(* IEC 61131-3 sources: plc-st-coding-agent/progress/evidence/f14_v14_remaining_20261113/jobs/codex_minimax-m27, 165 files *)

(* ---- public-easy-01.candidate_01.st ---- *)
(* ENGINEERING_CONTRACT *)
(*
  State machine for bottle filling line with 6 sequential states:
  - IDLE (0): No outputs active. Waits for bottleSensor TRUE → CLEANING.
  - CLEANING (1): Pump_Motor active. cleaningConfirmButton TRUE → FILLING.
  - FILLING (2): Filling_Valve active. fillingConfirmButton TRUE → CAPPING.
  - CAPPING (3): Capping_Machine active. cappingConfirmButton TRUE → PACKAGING.
  - PACKAGING (4): Packing_Machine active. packingConfirmButton TRUE → COMPLETED.
  - COMPLETED (5): Completion_Light active (retention). finishedButton TRUE → IDLE.

  Outputs: Pump_Motor(FILLING), Filling_Valve(FILLING), Capping_Machine(CAPPING),
           Packing_Machine(PACKAGING), Completion_Light(COMPLETED,hold_until_reset).
  Reset: finishedButton deactivates Completion_Light and returns to IDLE.
*)
(* CONTRACT_RULES [* kind=hold_until_reset, output=Completion_Light, set_input=packingConfirmButton, reset_input=finishedButton *] *)

FUNCTION_BLOCK FillingLineControl
VAR
    currentState : INT := 0;
END_VAR

CASE currentState OF
    0: // IDLE
        Pump_Motor := FALSE;
        Filling_Valve := FALSE;
        Capping_Machine := FALSE;
        Packing_Machine := FALSE;
        Completion_Light := FALSE;

        IF bottleSensor THEN
            currentState := 1;
        END_IF;

    1: // CLEANING
        Pump_Motor := TRUE;
        Filling_Valve := FALSE;
        Capping_Machine := FALSE;
        Packing_Machine := FALSE;
        Completion_Light := FALSE;

        IF cleaningConfirmButton THEN
            currentState := 2;
        END_IF;

    2: // FILLING
        Pump_Motor := FALSE;
        Filling_Valve := TRUE;
        Capping_Machine := FALSE;
        Packing_Machine := FALSE;
        Completion_Light := FALSE;

        IF fillingConfirmButton THEN
            currentState := 3;
        END_IF;

    3: // CAPPING
        Pump_Motor := FALSE;
        Filling_Valve := FALSE;
        Capping_Machine := TRUE;
        Packing_Machine := FALSE;
        Completion_Light := FALSE;

        IF cappingConfirmButton THEN
            currentState := 4;
        END_IF;

    4: // PACKAGING
        Pump_Motor := FALSE;
        Filling_Valve := FALSE;
        Capping_Machine := FALSE;
        Packing_Machine := TRUE;
        Completion_Light := FALSE;

        IF packingConfirmButton THEN
            currentState := 5;
        END_IF;

    5: // COMPLETED
        Pump_Motor := FALSE;
        Filling_Valve := FALSE;
        Capping_Machine := FALSE;
        Packing_Machine := FALSE;
        Completion_Light := TRUE;

        IF finishedButton THEN
            currentState := 0;
        END_IF;
END_CASE;
END_FUNCTION_BLOCK

(* ---- public-easy-01.candidate_03.st ---- *)
(* ENGINEERING_CONTRACT *)
(*
  State machine for bottle filling line with 6 sequential states:
  - IDLE (0): No outputs active. Waits for bottleSensor TRUE → CLEANING.
  - CLEANING (1): Pump_Motor active. cleaningConfirmButton TRUE → FILLING.
  - FILLING (2): Filling_Valve active. fillingConfirmButton TRUE → CAPPING.
  - CAPPING (3): Capping_Machine active. cappingConfirmButton TRUE → PACKAGING.
  - PACKAGING (4): Packing_Machine active. packingConfirmButton TRUE → COMPLETED.
  - COMPLETED (5): Completion_Light active (retention). finishedButton TRUE → IDLE.

  Outputs: Pump_Motor(FILLING), Filling_Valve(FILLING), Capping_Machine(CAPPING),
           Packing_Machine(PACKAGING), Completion_Light(COMPLETED,hold_until_reset).
  Reset: finishedButton deactivates Completion_Light and returns to IDLE.
*)
(* CONTRACT_RULES [* kind=hold_until_reset, output=Completion_Light, set_input=packingConfirmButton, reset_input=finishedButton *] *)

FUNCTION_BLOCK FillingLineControl
VAR_INPUT
    bottleSensor : BOOL;
    cleaningConfirmButton : BOOL;
    fillingConfirmButton : BOOL;
    cappingConfirmButton : BOOL;
    packingConfirmButton : BOOL;
    finishedButton : BOOL;
END_VAR
VAR_OUTPUT
    Pump_Motor : BOOL;
    Filling_Valve : BOOL;
    Capping_Machine : BOOL;
    Packing_Machine : BOOL;
    Completion_Light : BOOL;
END_VAR
VAR
    currentState : INT := 0;
END_VAR

CASE currentState OF
    0: // IDLE
        Pump_Motor := FALSE;
        Filling_Valve := FALSE;
        Capping_Machine := FALSE;
        Packing_Machine := FALSE;
        Completion_Light := FALSE;

        IF bottleSensor THEN
            currentState := 1;
        END_IF;

    1: // CLEANING
        Pump_Motor := TRUE;
        Filling_Valve := FALSE;
        Capping_Machine := FALSE;
        Packing_Machine := FALSE;
        Completion_Light := FALSE;

        IF cleaningConfirmButton THEN
            currentState := 2;
        END_IF;

    2: // FILLING
        Pump_Motor := FALSE;
        Filling_Valve := TRUE;
        Capping_Machine := FALSE;
        Packing_Machine := FALSE;
        Completion_Light := FALSE;

        IF fillingConfirmButton THEN
            currentState := 3;
        END_IF;

    3: // CAPPING
        Pump_Motor := FALSE;
        Filling_Valve := FALSE;
        Capping_Machine := TRUE;
        Packing_Machine := FALSE;
        Completion_Light := FALSE;

        IF cappingConfirmButton THEN
            currentState := 4;
        END_IF;

    4: // PACKAGING
        Pump_Motor := FALSE;
        Filling_Valve := FALSE;
        Capping_Machine := FALSE;
        Packing_Machine := TRUE;
        Completion_Light := FALSE;

        IF packingConfirmButton THEN
            currentState := 5;
        END_IF;

    5: // COMPLETED
        Pump_Motor := FALSE;
        Filling_Valve := FALSE;
        Capping_Machine := FALSE;
        Packing_Machine := FALSE;
        Completion_Light := TRUE;

        IF finishedButton THEN
            currentState := 0;
        END_IF;
END_CASE;
END_FUNCTION_BLOCK

(* ---- public-easy-01.patch_base_02.st ---- *)
(* ENGINEERING_CONTRACT *)
(*
  State machine for bottle filling line with 6 sequential states:
  - IDLE (0): No outputs active. Waits for bottleSensor TRUE → CLEANING.
  - CLEANING (1): Pump_Motor active. cleaningConfirmButton TRUE → FILLING.
  - FILLING (2): Filling_Valve active. fillingConfirmButton TRUE → CAPPING.
  - CAPPING (3): Capping_Machine active. cappingConfirmButton TRUE → PACKAGING.
  - PACKAGING (4): Packing_Machine active. packingConfirmButton TRUE → COMPLETED.
  - COMPLETED (5): Completion_Light active (retention). finishedButton TRUE → IDLE.

  Outputs: Pump_Motor(FILLING), Filling_Valve(FILLING), Capping_Machine(CAPPING),
           Packing_Machine(PACKAGING), Completion_Light(COMPLETED,hold_until_reset).
  Reset: finishedButton deactivates Completion_Light and returns to IDLE.
*)
(* CONTRACT_RULES [* kind=hold_until_reset, output=Completion_Light, set_input=packingConfirmButton, reset_input=finishedButton *] *)

FUNCTION_BLOCK FillingLineControl
VAR
    currentState : INT := 0;
END_VAR

CASE currentState OF
    0: // IDLE
        Pump_Motor := FALSE;
        Filling_Valve := FALSE;
        Capping_Machine := FALSE;
        Packing_Machine := FALSE;
        Completion_Light := FALSE;

        IF bottleSensor THEN
            currentState := 1;
        END_IF;

    1: // CLEANING
        Pump_Motor := TRUE;
        Filling_Valve := FALSE;
        Capping_Machine := FALSE;
        Packing_Machine := FALSE;
        Completion_Light := FALSE;

        IF cleaningConfirmButton THEN
            currentState := 2;
        END_IF;

    2: // FILLING
        Pump_Motor := FALSE;
        Filling_Valve := TRUE;
        Capping_Machine := FALSE;
        Packing_Machine := FALSE;
        Completion_Light := FALSE;

        IF fillingConfirmButton THEN
            currentState := 3;
        END_IF;

    3: // CAPPING
        Pump_Motor := FALSE;
        Filling_Valve := FALSE;
        Capping_Machine := TRUE;
        Packing_Machine := FALSE;
        Completion_Light := FALSE;

        IF cappingConfirmButton THEN
            currentState := 4;
        END_IF;

    4: // PACKAGING
        Pump_Motor := FALSE;
        Filling_Valve := FALSE;
        Capping_Machine := FALSE;
        Packing_Machine := TRUE;
        Completion_Light := FALSE;

        IF packingConfirmButton THEN
            currentState := 5;
        END_IF;

    5: // COMPLETED
        Pump_Motor := FALSE;
        Filling_Valve := FALSE;
        Capping_Machine := FALSE;
        Packing_Machine := FALSE;
        Completion_Light := TRUE;

        IF finishedButton THEN
            currentState := 0;
        END_IF;
END_CASE;
END_FUNCTION_BLOCK

(* ---- public-easy-01.patch_base_03.st ---- *)
(* ENGINEERING_CONTRACT *)
(*
  State machine for bottle filling line with 6 sequential states:
  - IDLE (0): No outputs active. Waits for bottleSensor TRUE → CLEANING.
  - CLEANING (1): Pump_Motor active. cleaningConfirmButton TRUE → FILLING.
  - FILLING (2): Filling_Valve active. fillingConfirmButton TRUE → CAPPING.
  - CAPPING (3): Capping_Machine active. cappingConfirmButton TRUE → PACKAGING.
  - PACKAGING (4): Packing_Machine active. packingConfirmButton TRUE → COMPLETED.
  - COMPLETED (5): Completion_Light active (retention). finishedButton TRUE → IDLE.

  Outputs: Pump_Motor(FILLING), Filling_Valve(FILLING), Capping_Machine(CAPPING),
           Packing_Machine(PACKAGING), Completion_Light(COMPLETED,hold_until_reset).
  Reset: finishedButton deactivates Completion_Light and returns to IDLE.
*)
(* CONTRACT_RULES [* kind=hold_until_reset, output=Completion_Light, set_input=packingConfirmButton, reset_input=finishedButton *] *)

FUNCTION_BLOCK FillingLineControl
VAR
    currentState : INT := 0;
END_VAR

CASE currentState OF
    0: // IDLE
        Pump_Motor := FALSE;
        Filling_Valve := FALSE;
        Capping_Machine := FALSE;
        Packing_Machine := FALSE;
        Completion_Light := FALSE;

        IF bottleSensor THEN
            currentState := 1;
        END_IF;

    1: // CLEANING
        Pump_Motor := TRUE;
        Filling_Valve := FALSE;
        Capping_Machine := FALSE;
        Packing_Machine := FALSE;
        Completion_Light := FALSE;

        IF cleaningConfirmButton THEN
            currentState := 2;
        END_IF;

    2: // FILLING
        Pump_Motor := FALSE;
        Filling_Valve := TRUE;
        Capping_Machine := FALSE;
        Packing_Machine := FALSE;
        Completion_Light := FALSE;

        IF fillingConfirmButton THEN
            currentState := 3;
        END_IF;

    3: // CAPPING
        Pump_Motor := FALSE;
        Filling_Valve := FALSE;
        Capping_Machine := TRUE;
        Packing_Machine := FALSE;
        Completion_Light := FALSE;

        IF cappingConfirmButton THEN
            currentState := 4;
        END_IF;

    4: // PACKAGING
        Pump_Motor := FALSE;
        Filling_Valve := FALSE;
        Capping_Machine := FALSE;
        Packing_Machine := TRUE;
        Completion_Light := FALSE;

        IF packingConfirmButton THEN
            currentState := 5;
        END_IF;

    5: // COMPLETED
        Pump_Motor := FALSE;
        Filling_Valve := FALSE;
        Capping_Machine := FALSE;
        Packing_Machine := FALSE;
        Completion_Light := TRUE;

        IF finishedButton THEN
            currentState := 0;
        END_IF;
END_CASE;
END_FUNCTION_BLOCK

(* ---- public-easy-01.patch_base_04.st ---- *)
(* ENGINEERING_CONTRACT *)
(*
  State machine for bottle filling line with 6 sequential states:
  - IDLE (0): No outputs active. Waits for bottleSensor TRUE → CLEANING.
  - CLEANING (1): Pump_Motor active. cleaningConfirmButton TRUE → FILLING.
  - FILLING (2): Filling_Valve active. fillingConfirmButton TRUE → CAPPING.
  - CAPPING (3): Capping_Machine active. cappingConfirmButton TRUE → PACKAGING.
  - PACKAGING (4): Packing_Machine active. packingConfirmButton TRUE → COMPLETED.
  - COMPLETED (5): Completion_Light active (retention). finishedButton TRUE → IDLE.

  Outputs: Pump_Motor(FILLING), Filling_Valve(FILLING), Capping_Machine(CAPPING),
           Packing_Machine(PACKAGING), Completion_Light(COMPLETED,hold_until_reset).
  Reset: finishedButton deactivates Completion_Light and returns to IDLE.
*)
(* CONTRACT_RULES [* kind=hold_until_reset, output=Completion_Light, set_input=packingConfirmButton, reset_input=finishedButton *] *)

FUNCTION_BLOCK FillingLineControl
VAR_INPUT
    bottleSensor : BOOL;
    cleaningConfirmButton : BOOL;
    fillingConfirmButton : BOOL;
    cappingConfirmButton : BOOL;
    packingConfirmButton : BOOL;
    finishedButton : BOOL;
END_VAR
VAR_OUTPUT
    Pump_Motor : BOOL;
    Filling_Valve : BOOL;
    Capping_Machine : BOOL;
    Packing_Machine : BOOL;
    Completion_Light : BOOL;
END_VAR
VAR
    currentState : INT := 0;
END_VAR

CASE currentState OF
    0: // IDLE
        Pump_Motor := FALSE;
        Filling_Valve := FALSE;
        Capping_Machine := FALSE;
        Packing_Machine := FALSE;
        Completion_Light := FALSE;

        IF bottleSensor THEN
            currentState := 1;
        END_IF;

    1: // CLEANING
        Pump_Motor := TRUE;
        Filling_Valve := FALSE;
        Capping_Machine := FALSE;
        Packing_Machine := FALSE;
        Completion_Light := FALSE;

        IF cleaningConfirmButton THEN
            currentState := 2;
        END_IF;

    2: // FILLING
        Pump_Motor := FALSE;
        Filling_Valve := TRUE;
        Capping_Machine := FALSE;
        Packing_Machine := FALSE;
        Completion_Light := FALSE;

        IF fillingConfirmButton THEN
            currentState := 3;
        END_IF;

    3: // CAPPING
        Pump_Motor := FALSE;
        Filling_Valve := FALSE;
        Capping_Machine := TRUE;
        Packing_Machine := FALSE;
        Completion_Light := FALSE;

        IF cappingConfirmButton THEN
            currentState := 4;
        END_IF;

    4: // PACKAGING
        Pump_Motor := FALSE;
        Filling_Valve := FALSE;
        Capping_Machine := FALSE;
        Packing_Machine := TRUE;
        Completion_Light := FALSE;

        IF packingConfirmButton THEN
            currentState := 5;
        END_IF;

    5: // COMPLETED
        Pump_Motor := FALSE;
        Filling_Valve := FALSE;
        Capping_Machine := FALSE;
        Packing_Machine := FALSE;
        Completion_Light := TRUE;

        IF finishedButton THEN
            currentState := 0;
        END_IF;
END_CASE;
END_FUNCTION_BLOCK

(* ---- public-easy-01.raw_candidate_01.st ---- *)
(* ENGINEERING_CONTRACT *)
(*
  State machine for bottle filling line with 6 sequential states:
  - IDLE (0): No outputs active. Waits for bottleSensor TRUE → CLEANING.
  - CLEANING (1): Pump_Motor active. cleaningConfirmButton TRUE → FILLING.
  - FILLING (2): Filling_Valve active. fillingConfirmButton TRUE → CAPPING.
  - CAPPING (3): Capping_Machine active. cappingConfirmButton TRUE → PACKAGING.
  - PACKAGING (4): Packing_Machine active. packingConfirmButton TRUE → COMPLETED.
  - COMPLETED (5): Completion_Light active (retention). finishedButton TRUE → IDLE.

  Outputs: Pump_Motor(FILLING), Filling_Valve(FILLING), Capping_Machine(CAPPING),
           Packing_Machine(PACKAGING), Completion_Light(COMPLETED,hold_until_reset).
  Reset: finishedButton deactivates Completion_Light and returns to IDLE.
*)
(* CONTRACT_RULES [* kind=hold_until_reset, output=Completion_Light, set_input=packingConfirmButton, reset_input=finishedButton *] *)

FUNCTION_BLOCK FillingLineControl
VAR
    currentState : INT := 0;
END_VAR

CASE currentState OF
    0: // IDLE
        Pump_Motor := FALSE;
        Filling_Valve := FALSE;
        Capping_Machine := FALSE;
        Packing_Machine := FALSE;
        Completion_Light := FALSE;

        IF bottleSensor THEN
            currentState := 1;
        END_IF;

    1: // CLEANING
        Pump_Motor := TRUE;
        Filling_Valve := FALSE;
        Capping_Machine := FALSE;
        Packing_Machine := FALSE;
        Completion_Light := FALSE;

        IF cleaningConfirmButton THEN
            currentState := 2;
        END_IF;

    2: // FILLING
        Pump_Motor := FALSE;
        Filling_Valve := TRUE;
        Capping_Machine := FALSE;
        Packing_Machine := FALSE;
        Completion_Light := FALSE;

        IF fillingConfirmButton THEN
            currentState := 3;
        END_IF;

    3: // CAPPING
        Pump_Motor := FALSE;
        Filling_Valve := FALSE;
        Capping_Machine := TRUE;
        Packing_Machine := FALSE;
        Completion_Light := FALSE;

        IF cappingConfirmButton THEN
            currentState := 4;
        END_IF;

    4: // PACKAGING
        Pump_Motor := FALSE;
        Filling_Valve := FALSE;
        Capping_Machine := FALSE;
        Packing_Machine := TRUE;
        Completion_Light := FALSE;

        IF packingConfirmButton THEN
            currentState := 5;
        END_IF;

    5: // COMPLETED
        Pump_Motor := FALSE;
        Filling_Valve := FALSE;
        Capping_Machine := FALSE;
        Packing_Machine := FALSE;
        Completion_Light := TRUE;

        IF finishedButton THEN
            currentState := 0;
        END_IF;
END_CASE;
END_FUNCTION_BLOCK

(* ---- public-easy-01.raw_candidate_03.st ---- *)
(* ENGINEERING_CONTRACT *)
(*
  State machine for bottle filling line with 6 sequential states:
  - IDLE (0): No outputs active. Waits for bottleSensor TRUE → CLEANING.
  - CLEANING (1): Pump_Motor active. cleaningConfirmButton TRUE → FILLING.
  - FILLING (2): Filling_Valve active. fillingConfirmButton TRUE → CAPPING.
  - CAPPING (3): Capping_Machine active. cappingConfirmButton TRUE → PACKAGING.
  - PACKAGING (4): Packing_Machine active. packingConfirmButton TRUE → COMPLETED.
  - COMPLETED (5): Completion_Light active (retention). finishedButton TRUE → IDLE.

  Outputs: Pump_Motor(FILLING), Filling_Valve(FILLING), Capping_Machine(CAPPING),
           Packing_Machine(PACKAGING), Completion_Light(COMPLETED,hold_until_reset).
  Reset: finishedButton deactivates Completion_Light and returns to IDLE.
*)
(* CONTRACT_RULES [* kind=hold_until_reset, output=Completion_Light, set_input=packingConfirmButton, reset_input=finishedButton *] *)

FUNCTION_BLOCK FillingLineControl
VAR_INPUT
    bottleSensor : BOOL;
    cleaningConfirmButton : BOOL;
    fillingConfirmButton : BOOL;
    cappingConfirmButton : BOOL;
    packingConfirmButton : BOOL;
    finishedButton : BOOL;
END_VAR
VAR_OUTPUT
    Pump_Motor : BOOL;
    Filling_Valve : BOOL;
    Capping_Machine : BOOL;
    Packing_Machine : BOOL;
    Completion_Light : BOOL;
END_VAR
VAR
    currentState : INT := 0;
END_VAR

CASE currentState OF
    0: // IDLE
        Pump_Motor := FALSE;
        Filling_Valve := FALSE;
        Capping_Machine := FALSE;
        Packing_Machine := FALSE;
        Completion_Light := FALSE;

        IF bottleSensor THEN
            currentState := 1;
        END_IF;

    1: // CLEANING
        Pump_Motor := TRUE;
        Filling_Valve := FALSE;
        Capping_Machine := FALSE;
        Packing_Machine := FALSE;
        Completion_Light := FALSE;

        IF cleaningConfirmButton THEN
            currentState := 2;
        END_IF;

    2: // FILLING
        Pump_Motor := FALSE;
        Filling_Valve := TRUE;
        Capping_Machine := FALSE;
        Packing_Machine := FALSE;
        Completion_Light := FALSE;

        IF fillingConfirmButton THEN
            currentState := 3;
        END_IF;

    3: // CAPPING
        Pump_Motor := FALSE;
        Filling_Valve := FALSE;
        Capping_Machine := TRUE;
        Packing_Machine := FALSE;
        Completion_Light := FALSE;

        IF cappingConfirmButton THEN
            currentState := 4;
        END_IF;

    4: // PACKAGING
        Pump_Motor := FALSE;
        Filling_Valve := FALSE;
        Capping_Machine := FALSE;
        Packing_Machine := TRUE;
        Completion_Light := FALSE;

        IF packingConfirmButton THEN
            currentState := 5;
        END_IF;

    5: // COMPLETED
        Pump_Motor := FALSE;
        Filling_Valve := FALSE;
        Capping_Machine := FALSE;
        Packing_Machine := FALSE;
        Completion_Light := TRUE;

        IF finishedButton THEN
            currentState := 0;
        END_IF;
END_CASE;
END_FUNCTION_BLOCK

(* ---- public-easy-02.candidate_01.st ---- *)
FUNCTION_BLOCK FB_DualWordEdgeDetection
VAR_INPUT
    value : DWORD;
END_VAR
VAR_OUTPUT
    hasChanged     : BOOL;
    hasRisingEdges : BOOL;
    risingBits     : DWORD;
    noOfRisingBits : USINT;
    hasFallingEdges: BOOL;
    fallingBits    : DWORD;
    noOfFallingBits: USINT;
END_VAR
VAR
    prevValue : DWORD;
END_VAR

(*
ENGINEERING_CONTRACT
==================
PUB001: Edge detection per bit of DWORD input, all 32 bits tracked independently
Activation:    Continuous, outputs update every scan cycle
Retention:     prevValue retains last cycle state; risingBits/fallingBits valid for current scan only
Reset/Deact:   No explicit reset input - prevValue updates automatically each cycle
Same-scan:     Uses prevValue from previous invocation for edge calculation
Units:         BIT positions 0-31; counts are 0-32
Boundary:      32-bit DWORD; all operations use DWORD arithmetic
==================
*)

risingBits  := value AND (NOT prevValue);
fallingBits := (NOT value) AND prevValue;

hasChanged     := (value <> prevValue);
hasRisingEdges := (risingBits <> 16#0);
hasFallingEdges:= (fallingBits <> 16#0);

noOfRisingBits  := TO_USINT(SHL(value, 24) <> 16#0) + TO_USINT(SHL(value, 25) <> 16#0) +
                   TO_USINT(SHL(value, 26) <> 16#0) + TO_USINT(SHL(value, 27) <> 16#0) +
                   TO_USINT(SHL(value, 28) <> 16#0) + TO_USINT(SHL(value, 29) <> 16#0) +
                   TO_USINT(SHL(value, 30) <> 16#0) + TO_USINT(SHL(value, 31) <> 16#0);

noOfFallingBits := TO_USINT(SHL(fallingBits, 24) <> 16#0) + TO_USINT(SHL(fallingBits, 25) <> 16#0) +
                   TO_USINT(SHL(fallingBits, 26) <> 16#0) + TO_USINT(SHL(fallingBits, 27) <> 16#0) +
                   TO_USINT(SHL(fallingBits, 28) <> 16#0) + TO_USINT(SHL(fallingBits, 29) <> 16#0) +
                   TO_USINT(SHL(fallingBits, 30) <> 16#0) + TO_USINT(SHL(fallingBits, 31) <> 16#0);

prevValue := value;
END_FUNCTION_BLOCK

(* ---- public-easy-02.candidate_03.st ---- *)
FUNCTION_BLOCK FB_DualWordEdgeDetection
VAR_INPUT
    value : DWORD;
END_VAR
VAR_OUTPUT
    hasChanged     : BOOL;
    hasRisingEdges : BOOL;
    risingBits     : DWORD;
    noOfRisingBits : USINT;
    hasFallingEdges: BOOL;
    fallingBits    : DWORD;
    noOfFallingBits: USINT;
END_VAR
VAR
    prevValue : DWORD;
END_VAR

(*
ENGINEERING_CONTRACT
==================
PUB001: Edge detection per bit of DWORD input, all 32 bits tracked independently
Activation:    Continuous, outputs update every scan cycle
Retention:     prevValue retains last cycle state; risingBits/fallingBits valid for current scan only
Reset/Deact:   No explicit reset input - prevValue updates automatically each cycle
Same-scan:     Uses prevValue from previous invocation for edge calculation
Units:         BIT positions 0-31; counts are 0-32
Boundary:      32-bit DWORD; all operations use DWORD arithmetic
==================
*)

risingBits  := value AND (NOT prevValue);
fallingBits := (NOT value) AND prevValue;

hasChanged     := (value <> prevValue);
hasRisingEdges := (risingBits <> 16#0);
hasFallingEdges:= (fallingBits <> 16#0);

noOfRisingBits  := 0;
FOR tmp_i := 0 TO 31 DO
    IF (risingBits SHR TO_USINT(tmp_i)) AND 16#1 = 1 THEN
        noOfRisingBits := noOfRisingBits + 1;
    END_IF;
END_FOR;

noOfFallingBits := 0;
FOR tmp_i := 0 TO 31 DO
    IF (fallingBits SHR TO_USINT(tmp_i)) AND 16#1 = 1 THEN
        noOfFallingBits := noOfFallingBits + 1;
    END_IF;
END_FOR;

prevValue := value;
END_FUNCTION_BLOCK

(* ---- public-easy-02.patch_base_02.st ---- *)
FUNCTION_BLOCK FB_DualWordEdgeDetection
VAR_INPUT
    value : DWORD;
END_VAR
VAR_OUTPUT
    hasChanged     : BOOL;
    hasRisingEdges : BOOL;
    risingBits     : DWORD;
    noOfRisingBits : USINT;
    hasFallingEdges: BOOL;
    fallingBits    : DWORD;
    noOfFallingBits: USINT;
END_VAR
VAR
    prevValue : DWORD;
END_VAR

(*
ENGINEERING_CONTRACT
==================
PUB001: Edge detection per bit of DWORD input, all 32 bits tracked independently
Activation:    Continuous, outputs update every scan cycle
Retention:     prevValue retains last cycle state; risingBits/fallingBits valid for current scan only
Reset/Deact:   No explicit reset input - prevValue updates automatically each cycle
Same-scan:     Uses prevValue from previous invocation for edge calculation
Units:         BIT positions 0-31; counts are 0-32
Boundary:      32-bit DWORD; all operations use DWORD arithmetic
==================
*)

risingBits  := value AND (NOT prevValue);
fallingBits := (NOT value) AND prevValue;

hasChanged     := (value <> prevValue);
hasRisingEdges := (risingBits <> 16#0);
hasFallingEdges:= (fallingBits <> 16#0);

noOfRisingBits  := TO_USINT(SHL(value, 24) <> 16#0) + TO_USINT(SHL(value, 25) <> 16#0) +
                   TO_USINT(SHL(value, 26) <> 16#0) + TO_USINT(SHL(value, 27) <> 16#0) +
                   TO_USINT(SHL(value, 28) <> 16#0) + TO_USINT(SHL(value, 29) <> 16#0) +
                   TO_USINT(SHL(value, 30) <> 16#0) + TO_USINT(SHL(value, 31) <> 16#0);

noOfFallingBits := TO_USINT(SHL(fallingBits, 24) <> 16#0) + TO_USINT(SHL(fallingBits, 25) <> 16#0) +
                   TO_USINT(SHL(fallingBits, 26) <> 16#0) + TO_USINT(SHL(fallingBits, 27) <> 16#0) +
                   TO_USINT(SHL(fallingBits, 28) <> 16#0) + TO_USINT(SHL(fallingBits, 29) <> 16#0) +
                   TO_USINT(SHL(fallingBits, 30) <> 16#0) + TO_USINT(SHL(fallingBits, 31) <> 16#0);

prevValue := value;
END_FUNCTION_BLOCK

(* ---- public-easy-02.patch_base_03.st ---- *)
FUNCTION_BLOCK FB_DualWordEdgeDetection
VAR_INPUT
    value : DWORD;
END_VAR
VAR_OUTPUT
    hasChanged     : BOOL;
    hasRisingEdges : BOOL;
    risingBits     : DWORD;
    noOfRisingBits : USINT;
    hasFallingEdges: BOOL;
    fallingBits    : DWORD;
    noOfFallingBits: USINT;
END_VAR
VAR
    prevValue : DWORD;
END_VAR

(*
ENGINEERING_CONTRACT
==================
PUB001: Edge detection per bit of DWORD input, all 32 bits tracked independently
Activation:    Continuous, outputs update every scan cycle
Retention:     prevValue retains last cycle state; risingBits/fallingBits valid for current scan only
Reset/Deact:   No explicit reset input - prevValue updates automatically each cycle
Same-scan:     Uses prevValue from previous invocation for edge calculation
Units:         BIT positions 0-31; counts are 0-32
Boundary:      32-bit DWORD; all operations use DWORD arithmetic
==================
*)

risingBits  := value AND (NOT prevValue);
fallingBits := (NOT value) AND prevValue;

hasChanged     := (value <> prevValue);
hasRisingEdges := (risingBits <> 16#0);
hasFallingEdges:= (fallingBits <> 16#0);

noOfRisingBits  := TO_USINT(SHL(value, 24) <> 16#0) + TO_USINT(SHL(value, 25) <> 16#0) +
                   TO_USINT(SHL(value, 26) <> 16#0) + TO_USINT(SHL(value, 27) <> 16#0) +
                   TO_USINT(SHL(value, 28) <> 16#0) + TO_USINT(SHL(value, 29) <> 16#0) +
                   TO_USINT(SHL(value, 30) <> 16#0) + TO_USINT(SHL(value, 31) <> 16#0);

noOfFallingBits := TO_USINT(SHL(fallingBits, 24) <> 16#0) + TO_USINT(SHL(fallingBits, 25) <> 16#0) +
                   TO_USINT(SHL(fallingBits, 26) <> 16#0) + TO_USINT(SHL(fallingBits, 27) <> 16#0) +
                   TO_USINT(SHL(fallingBits, 28) <> 16#0) + TO_USINT(SHL(fallingBits, 29) <> 16#0) +
                   TO_USINT(SHL(fallingBits, 30) <> 16#0) + TO_USINT(SHL(fallingBits, 31) <> 16#0);

prevValue := value;
END_FUNCTION_BLOCK

(* ---- public-easy-02.patch_base_04.st ---- *)
FUNCTION_BLOCK FB_DualWordEdgeDetection
VAR_INPUT
    value : DWORD;
END_VAR
VAR_OUTPUT
    hasChanged     : BOOL;
    hasRisingEdges : BOOL;
    risingBits     : DWORD;
    noOfRisingBits : USINT;
    hasFallingEdges: BOOL;
    fallingBits    : DWORD;
    noOfFallingBits: USINT;
END_VAR
VAR
    prevValue : DWORD;
END_VAR

(*
ENGINEERING_CONTRACT
==================
PUB001: Edge detection per bit of DWORD input, all 32 bits tracked independently
Activation:    Continuous, outputs update every scan cycle
Retention:     prevValue retains last cycle state; risingBits/fallingBits valid for current scan only
Reset/Deact:   No explicit reset input - prevValue updates automatically each cycle
Same-scan:     Uses prevValue from previous invocation for edge calculation
Units:         BIT positions 0-31; counts are 0-32
Boundary:      32-bit DWORD; all operations use DWORD arithmetic
==================
*)

risingBits  := value AND (NOT prevValue);
fallingBits := (NOT value) AND prevValue;

hasChanged     := (value <> prevValue);
hasRisingEdges := (risingBits <> 16#0);
hasFallingEdges:= (fallingBits <> 16#0);

noOfRisingBits  := TO_USINT(SHL(value, 24) <> 16#0) + TO_USINT(SHL(value, 25) <> 16#0) +
                   TO_USINT(SHL(value, 26) <> 16#0) + TO_USINT(SHL(value, 27) <> 16#0) +
                   TO_USINT(SHL(value, 28) <> 16#0) + TO_USINT(SHL(value, 29) <> 16#0) +
                   TO_USINT(SHL(value, 30) <> 16#0) + TO_USINT(SHL(value, 31) <> 16#0);

noOfFallingBits := TO_USINT(SHL(fallingBits, 24) <> 16#0) + TO_USINT(SHL(fallingBits, 25) <> 16#0) +
                   TO_USINT(SHL(fallingBits, 26) <> 16#0) + TO_USINT(SHL(fallingBits, 27) <> 16#0) +
                   TO_USINT(SHL(fallingBits, 28) <> 16#0) + TO_USINT(SHL(fallingBits, 29) <> 16#0) +
                   TO_USINT(SHL(fallingBits, 30) <> 16#0) + TO_USINT(SHL(fallingBits, 31) <> 16#0);

prevValue := value;
END_FUNCTION_BLOCK

(* ---- public-easy-02.raw_candidate_01.st ---- *)
FUNCTION_BLOCK FB_DualWordEdgeDetection
VAR_INPUT
    value : DWORD;
END_VAR
VAR_OUTPUT
    hasChanged     : BOOL;
    hasRisingEdges : BOOL;
    risingBits     : DWORD;
    noOfRisingBits : USINT;
    hasFallingEdges: BOOL;
    fallingBits    : DWORD;
    noOfFallingBits: USINT;
END_VAR
VAR
    prevValue : DWORD;
END_VAR

(*
ENGINEERING_CONTRACT
==================
PUB001: Edge detection per bit of DWORD input, all 32 bits tracked independently
Activation:    Continuous, outputs update every scan cycle
Retention:     prevValue retains last cycle state; risingBits/fallingBits valid for current scan only
Reset/Deact:   No explicit reset input - prevValue updates automatically each cycle
Same-scan:     Uses prevValue from previous invocation for edge calculation
Units:         BIT positions 0-31; counts are 0-32
Boundary:      32-bit DWORD; all operations use DWORD arithmetic
==================
*)

risingBits  := value AND (NOT prevValue);
fallingBits := (NOT value) AND prevValue;

hasChanged     := (value <> prevValue);
hasRisingEdges := (risingBits <> 16#0);
hasFallingEdges:= (fallingBits <> 16#0);

noOfRisingBits  := TO_USINT(SHL(value, 24) <> 16#0) + TO_USINT(SHL(value, 25) <> 16#0) +
                   TO_USINT(SHL(value, 26) <> 16#0) + TO_USINT(SHL(value, 27) <> 16#0) +
                   TO_USINT(SHL(value, 28) <> 16#0) + TO_USINT(SHL(value, 29) <> 16#0) +
                   TO_USINT(SHL(value, 30) <> 16#0) + TO_USINT(SHL(value, 31) <> 16#0);

noOfFallingBits := TO_USINT(SHL(fallingBits, 24) <> 16#0) + TO_USINT(SHL(fallingBits, 25) <> 16#0) +
                   TO_USINT(SHL(fallingBits, 26) <> 16#0) + TO_USINT(SHL(fallingBits, 27) <> 16#0) +
                   TO_USINT(SHL(fallingBits, 28) <> 16#0) + TO_USINT(SHL(fallingBits, 29) <> 16#0) +
                   TO_USINT(SHL(fallingBits, 30) <> 16#0) + TO_USINT(SHL(fallingBits, 31) <> 16#0);

prevValue := value;
END_FUNCTION_BLOCK

(* ---- public-easy-02.raw_candidate_03.st ---- *)
FUNCTION_BLOCK FB_DualWordEdgeDetection
VAR_INPUT
    value : DWORD;
END_VAR
VAR_OUTPUT
    hasChanged     : BOOL;
    hasRisingEdges : BOOL;
    risingBits     : DWORD;
    noOfRisingBits : USINT;
    hasFallingEdges: BOOL;
    fallingBits    : DWORD;
    noOfFallingBits: USINT;
END_VAR
VAR
    prevValue : DWORD;
END_VAR

(*
ENGINEERING_CONTRACT
==================
PUB001: Edge detection per bit of DWORD input, all 32 bits tracked independently
Activation:    Continuous, outputs update every scan cycle
Retention:     prevValue retains last cycle state; risingBits/fallingBits valid for current scan only
Reset/Deact:   No explicit reset input - prevValue updates automatically each cycle
Same-scan:     Uses prevValue from previous invocation for edge calculation
Units:         BIT positions 0-31; counts are 0-32
Boundary:      32-bit DWORD; all operations use DWORD arithmetic
==================
*)

risingBits  := value AND (NOT prevValue);
fallingBits := (NOT value) AND prevValue;

hasChanged     := (value <> prevValue);
hasRisingEdges := (risingBits <> 16#0);
hasFallingEdges:= (fallingBits <> 16#0);

noOfRisingBits  := 0;
FOR tmp_i := 0 TO 31 DO
    IF (risingBits SHR TO_USINT(tmp_i)) AND 16#1 = 1 THEN
        noOfRisingBits := noOfRisingBits + 1;
    END_IF;
END_FOR;

noOfFallingBits := 0;
FOR tmp_i := 0 TO 31 DO
    IF (fallingBits SHR TO_USINT(tmp_i)) AND 16#1 = 1 THEN
        noOfFallingBits := noOfFallingBits + 1;
    END_IF;
END_FOR;

prevValue := value;
END_FUNCTION_BLOCK

(* ---- public-easy-03.candidate_01.st ---- *)
(*
ENGINEERING_CONTRACT
===================
hiAlarm activation: Value > hiLevel (PUB001)
hiAlarm retention: remains TRUE until Value < hiLevel - hystWindow (PUB001)
loAlarm activation: Value < loLevel (PUB003)
loAlarm retention: remains TRUE until Value > loLevel + hystWindow (PUB003)
error activation: loLevel >= hiLevel → status=16#8001 (PUB005)
error activation: hystWindow >= (hiLevel - loLevel) → status=16#8002 (PUB006)
reset/deactivation: error conditions return early, alarms retain prior state
same-scan priority: error checks precede alarm logic; no output overlap conflicts
units/boundaries: REAL comparisons with explicit thresholds; strict > and <

CONTRACT_RULES []
*)

FUNCTION_BLOCK AlarmHysteresis
VAR_INPUT
    Value       : REAL;
    hiLevel     : REAL;
    loLevel     : REAL;
    hystWindow  : REAL;
END_VAR
VAR_OUTPUT
    hiAlarm     : BOOL := FALSE;
    loAlarm     : BOOL := FALSE;
    error       : BOOL := FALSE;
    status      : WORD := 16#0000;
END_VAR
VAR
END_VAR

// Parameter validation: loLevel must be less than hiLevel
IF loLevel >= hiLevel THEN
    error := TRUE;
    status := 16#8001;
    RETURN;
END_IF;

// Parameter validation: hystWindow must be less than the range between hiLevel and loLevel
IF hystWindow >= (hiLevel - loLevel) THEN
    error := TRUE;
    status := 16#8002;
    RETURN;
END_IF;

// High alarm: trigger when Value exceeds hiLevel, clear when below hiLevel minus hysteresis
IF Value > hiLevel THEN
    hiAlarm := TRUE;
ELSIF Value < (hiLevel - hystWindow) THEN
    hiAlarm := FALSE;
END_IF;

// Low alarm: trigger when Value falls below loLevel, clear when above loLevel plus hysteresis
IF Value < loLevel THEN
    loAlarm := TRUE;
ELSIF Value > (loLevel + hystWindow) THEN
    loAlarm := FALSE;
END_IF;

END_FUNCTION_BLOCK

(* ---- public-easy-03.candidate_03.st ---- *)
(*
ENGINEERING_CONTRACT
===================
hiAlarm activation: Value > hiLevel (PUB001)
hiAlarm retention: remains TRUE until Value < hiLevel - hystWindow (PUB001)
loAlarm activation: Value < loLevel (PUB003)
loAlarm retention: remains TRUE until Value > loLevel + hystWindow (PUB003)
error activation: loLevel >= hiLevel → status=16#8001 (PUB005)
error activation: hystWindow >= (hiLevel - loLevel) → status=16#8002 (PUB006)
reset/deactivation: error conditions return early, alarms retain prior state
same-scan priority: error checks precede alarm logic; no output overlap conflicts
units/boundaries: REAL comparisons with explicit thresholds; strict > and <

CONTRACT_RULES []
*)

FUNCTION_BLOCK AlarmHysteresis
VAR_INPUT
    Value       : REAL;
    hiLevel     : REAL;
    loLevel     : REAL;
    hystWindow  : REAL;
END_VAR
VAR_OUTPUT
    hiAlarm     : BOOL := FALSE;
    loAlarm     : BOOL := FALSE;
    error       : BOOL := FALSE;
    status      : WORD := 16#0000;
END_VAR
VAR
    tmpError    : BOOL := FALSE;
    tmpStatus   : WORD := 16#0000;
END_VAR

IF loLevel >= hiLevel THEN
    tmpError := TRUE;
    tmpStatus := 16#8001;
END_IF;

IF hystWindow >= (hiLevel - loLevel) THEN
    tmpError := TRUE;
    tmpStatus := 16#8002;
END_IF;

error := tmpError;
status := tmpStatus;

IF NOT tmpError THEN
    IF Value > hiLevel THEN
        hiAlarm := TRUE;
    ELSIF Value < (hiLevel - hystWindow) THEN
        hiAlarm := FALSE;
    END_IF;

    IF Value < loLevel THEN
        loAlarm := TRUE;
    ELSIF Value > (loLevel + hystWindow) THEN
        loAlarm := FALSE;
    END_IF;
END_IF;

END_FUNCTION_BLOCK

(* ---- public-easy-03.patch_base_02.st ---- *)
(*
ENGINEERING_CONTRACT
===================
hiAlarm activation: Value > hiLevel (PUB001)
hiAlarm retention: remains TRUE until Value < hiLevel - hystWindow (PUB001)
loAlarm activation: Value < loLevel (PUB003)
loAlarm retention: remains TRUE until Value > loLevel + hystWindow (PUB003)
error activation: loLevel >= hiLevel → status=16#8001 (PUB005)
error activation: hystWindow >= (hiLevel - loLevel) → status=16#8002 (PUB006)
reset/deactivation: error conditions return early, alarms retain prior state
same-scan priority: error checks precede alarm logic; no output overlap conflicts
units/boundaries: REAL comparisons with explicit thresholds; strict > and <

CONTRACT_RULES []
*)

FUNCTION_BLOCK AlarmHysteresis
VAR_INPUT
    Value       : REAL;
    hiLevel     : REAL;
    loLevel     : REAL;
    hystWindow  : REAL;
END_VAR
VAR_OUTPUT
    hiAlarm     : BOOL := FALSE;
    loAlarm     : BOOL := FALSE;
    error       : BOOL := FALSE;
    status      : WORD := 16#0000;
END_VAR
VAR
END_VAR

// Parameter validation: loLevel must be less than hiLevel
IF loLevel >= hiLevel THEN
    error := TRUE;
    status := 16#8001;
    RETURN;
END_IF;

// Parameter validation: hystWindow must be less than the range between hiLevel and loLevel
IF hystWindow >= (hiLevel - loLevel) THEN
    error := TRUE;
    status := 16#8002;
    RETURN;
END_IF;

// High alarm: trigger when Value exceeds hiLevel, clear when below hiLevel minus hysteresis
IF Value > hiLevel THEN
    hiAlarm := TRUE;
ELSIF Value < (hiLevel - hystWindow) THEN
    hiAlarm := FALSE;
END_IF;

// Low alarm: trigger when Value falls below loLevel, clear when above loLevel plus hysteresis
IF Value < loLevel THEN
    loAlarm := TRUE;
ELSIF Value > (loLevel + hystWindow) THEN
    loAlarm := FALSE;
END_IF;

END_FUNCTION_BLOCK

(* ---- public-easy-03.patch_base_03.st ---- *)
(*
ENGINEERING_CONTRACT
===================
hiAlarm activation: Value > hiLevel (PUB001)
hiAlarm retention: remains TRUE until Value < hiLevel - hystWindow (PUB001)
loAlarm activation: Value < loLevel (PUB003)
loAlarm retention: remains TRUE until Value > loLevel + hystWindow (PUB003)
error activation: loLevel >= hiLevel → status=16#8001 (PUB005)
error activation: hystWindow >= (hiLevel - loLevel) → status=16#8002 (PUB006)
reset/deactivation: error conditions return early, alarms retain prior state
same-scan priority: error checks precede alarm logic; no output overlap conflicts
units/boundaries: REAL comparisons with explicit thresholds; strict > and <

CONTRACT_RULES []
*)

FUNCTION_BLOCK AlarmHysteresis
VAR_INPUT
    Value       : REAL;
    hiLevel     : REAL;
    loLevel     : REAL;
    hystWindow  : REAL;
END_VAR
VAR_OUTPUT
    hiAlarm     : BOOL := FALSE;
    loAlarm     : BOOL := FALSE;
    error       : BOOL := FALSE;
    status      : WORD := 16#0000;
END_VAR
VAR
END_VAR

// Parameter validation: loLevel must be less than hiLevel
IF loLevel >= hiLevel THEN
    error := TRUE;
    status := 16#8001;
    RETURN;
END_IF;

// Parameter validation: hystWindow must be less than the range between hiLevel and loLevel
IF hystWindow >= (hiLevel - loLevel) THEN
    error := TRUE;
    status := 16#8002;
    RETURN;
END_IF;

// High alarm: trigger when Value exceeds hiLevel, clear when below hiLevel minus hysteresis
IF Value > hiLevel THEN
    hiAlarm := TRUE;
ELSIF Value < (hiLevel - hystWindow) THEN
    hiAlarm := FALSE;
END_IF;

// Low alarm: trigger when Value falls below loLevel, clear when above loLevel plus hysteresis
IF Value < loLevel THEN
    loAlarm := TRUE;
ELSIF Value > (loLevel + hystWindow) THEN
    loAlarm := FALSE;
END_IF;

END_FUNCTION_BLOCK

(* ---- public-easy-03.patch_base_04.st ---- *)
(*
ENGINEERING_CONTRACT
===================
hiAlarm activation: Value > hiLevel (PUB001)
hiAlarm retention: remains TRUE until Value < hiLevel - hystWindow (PUB001)
loAlarm activation: Value < loLevel (PUB003)
loAlarm retention: remains TRUE until Value > loLevel + hystWindow (PUB003)
error activation: loLevel >= hiLevel → status=16#8001 (PUB005)
error activation: hystWindow >= (hiLevel - loLevel) → status=16#8002 (PUB006)
reset/deactivation: error conditions return early, alarms retain prior state
same-scan priority: error checks precede alarm logic; no output overlap conflicts
units/boundaries: REAL comparisons with explicit thresholds; strict > and <

CONTRACT_RULES []
*)

FUNCTION_BLOCK AlarmHysteresis
VAR_INPUT
    Value       : REAL;
    hiLevel     : REAL;
    loLevel     : REAL;
    hystWindow  : REAL;
END_VAR
VAR_OUTPUT
    hiAlarm     : BOOL := FALSE;
    loAlarm     : BOOL := FALSE;
    error       : BOOL := FALSE;
    status      : WORD := 16#0000;
END_VAR
VAR
END_VAR

// Parameter validation: loLevel must be less than hiLevel
IF loLevel >= hiLevel THEN
    error := TRUE;
    status := 16#8001;
    RETURN;
END_IF;

// Parameter validation: hystWindow must be less than the range between hiLevel and loLevel
IF hystWindow >= (hiLevel - loLevel) THEN
    error := TRUE;
    status := 16#8002;
    RETURN;
END_IF;

// High alarm: trigger when Value exceeds hiLevel, clear when below hiLevel minus hysteresis
IF Value > hiLevel THEN
    hiAlarm := TRUE;
ELSIF Value < (hiLevel - hystWindow) THEN
    hiAlarm := FALSE;
END_IF;

// Low alarm: trigger when Value falls below loLevel, clear when above loLevel plus hysteresis
IF Value < loLevel THEN
    loAlarm := TRUE;
ELSIF Value > (loLevel + hystWindow) THEN
    loAlarm := FALSE;
END_IF;

END_FUNCTION_BLOCK

(* ---- public-easy-03.raw_candidate_01.st ---- *)
(*
ENGINEERING_CONTRACT
===================
hiAlarm activation: Value > hiLevel (PUB001)
hiAlarm retention: remains TRUE until Value < hiLevel - hystWindow (PUB001)
loAlarm activation: Value < loLevel (PUB003)
loAlarm retention: remains TRUE until Value > loLevel + hystWindow (PUB003)
error activation: loLevel >= hiLevel → status=16#8001 (PUB005)
error activation: hystWindow >= (hiLevel - loLevel) → status=16#8002 (PUB006)
reset/deactivation: error conditions return early, alarms retain prior state
same-scan priority: error checks precede alarm logic; no output overlap conflicts
units/boundaries: REAL comparisons with explicit thresholds; strict > and <

CONTRACT_RULES []
*)

FUNCTION_BLOCK AlarmHysteresis
VAR_INPUT
    Value       : REAL;
    hiLevel     : REAL;
    loLevel     : REAL;
    hystWindow  : REAL;
END_VAR
VAR_OUTPUT
    hiAlarm     : BOOL := FALSE;
    loAlarm     : BOOL := FALSE;
    error       : BOOL := FALSE;
    status      : WORD := 16#0000;
END_VAR
VAR
END_VAR

// Parameter validation: loLevel must be less than hiLevel
IF loLevel >= hiLevel THEN
    error := TRUE;
    status := 16#8001;
    RETURN;
END_IF;

// Parameter validation: hystWindow must be less than the range between hiLevel and loLevel
IF hystWindow >= (hiLevel - loLevel) THEN
    error := TRUE;
    status := 16#8002;
    RETURN;
END_IF;

// High alarm: trigger when Value exceeds hiLevel, clear when below hiLevel minus hysteresis
IF Value > hiLevel THEN
    hiAlarm := TRUE;
ELSIF Value < (hiLevel - hystWindow) THEN
    hiAlarm := FALSE;
END_IF;

// Low alarm: trigger when Value falls below loLevel, clear when above loLevel plus hysteresis
IF Value < loLevel THEN
    loAlarm := TRUE;
ELSIF Value > (loLevel + hystWindow) THEN
    loAlarm := FALSE;
END_IF;

END_FUNCTION_BLOCK

(* ---- public-easy-03.raw_candidate_03.st ---- *)
(*
ENGINEERING_CONTRACT
===================
hiAlarm activation: Value > hiLevel (PUB001)
hiAlarm retention: remains TRUE until Value < hiLevel - hystWindow (PUB001)
loAlarm activation: Value < loLevel (PUB003)
loAlarm retention: remains TRUE until Value > loLevel + hystWindow (PUB003)
error activation: loLevel >= hiLevel → status=16#8001 (PUB005)
error activation: hystWindow >= (hiLevel - loLevel) → status=16#8002 (PUB006)
reset/deactivation: error conditions return early, alarms retain prior state
same-scan priority: error checks precede alarm logic; no output overlap conflicts
units/boundaries: REAL comparisons with explicit thresholds; strict > and <

CONTRACT_RULES []
*)

FUNCTION_BLOCK AlarmHysteresis
VAR_INPUT
    Value       : REAL;
    hiLevel     : REAL;
    loLevel     : REAL;
    hystWindow  : REAL;
END_VAR
VAR_OUTPUT
    hiAlarm     : BOOL := FALSE;
    loAlarm     : BOOL := FALSE;
    error       : BOOL := FALSE;
    status      : WORD := 16#0000;
END_VAR
VAR
    tmpError    : BOOL := FALSE;
    tmpStatus   : WORD := 16#0000;
END_VAR

IF loLevel >= hiLevel THEN
    tmpError := TRUE;
    tmpStatus := 16#8001;
END_IF;

IF hystWindow >= (hiLevel - loLevel) THEN
    tmpError := TRUE;
    tmpStatus := 16#8002;
END_IF;

error := tmpError;
status := tmpStatus;

IF NOT tmpError THEN
    IF Value > hiLevel THEN
        hiAlarm := TRUE;
    ELSIF Value < (hiLevel - hystWindow) THEN
        hiAlarm := FALSE;
    END_IF;

    IF Value < loLevel THEN
        loAlarm := TRUE;
    ELSIF Value > (loLevel + hystWindow) THEN
        loAlarm := FALSE;
    END_IF;
END_IF;

END_FUNCTION_BLOCK

(* ---- public-easy-04.candidate_01.st ---- *)
FUNCTION_BLOCK JamPumpControl
VAR_INPUT
    VISCOSITY_OK    : BOOL;
    PASTE_E_STOP_NC : BOOL;
    DebounceTime    : TIME;
    CycleTime       : TIME;
END_VAR

VAR_OUTPUT
    VFD_RUN          : BOOL := FALSE;
    PUMP_MAINT_DUE   : BOOL := FALSE;
    PUMP_RUNTIME_ACC : LTIME := LTIME#0s;
END_VAR

VAR
    viscosityTimer : TON;
    viscosityValid : BOOL := FALSE;
END_VAR

(* ENGINEERING_CONTRACT
 * =============================================================================
 * Output: VFD_RUN
 *   - Activation:   PASTE_E_STOP_NC = TRUE AND viscosityValid = TRUE (PUB001, PUB002)
 *   - Retention:    Held TRUE while both permissive conditions remain TRUE
 *   - Reset:        Immediate on PASTE_E_STOP_NC = FALSE (E-stop) OR viscosityValid = FALSE
 *   - Same-scan:    E-stop has highest priority; cleared first scan of E-stop event
 *   - Units:        Boolean command, no time units
 * ----------------------------------------------------------------------------
 * Output: PUMP_RUNTIME_ACC
 *   - Activation:   VFD_RUN = TRUE (PUB003)
 *   - Retention:    Preserved while VFD_RUN = FALSE; never cleared by E-stop
 *   - Reset:        None (informational only)
 *   - Same-scan:    Accumulates once per invocation using CycleTime value
 *   - Units:        LTIME nanoseconds; 500h = 1,800,000,000,000 ns (PUB004)
 * ----------------------------------------------------------------------------
 * Output: PUMP_MAINT_DUE
 *   - Activation:   PUMP_RUNTIME_ACC >= 500 hours (PUB004)
 *   - Retention:    Held TRUE once threshold reached (no explicit reset required)
 *   - Reset:        None stated; informational only
 *   - Same-scan:    Evaluated every invocation
 *   - Units:        Boolean indication, does not affect VFD_RUN or safety permissive
 * ----------------------------------------------------------------------------
 * Internal: viscosityValid
 *   - Activation:   VISCOSITY_OK = TRUE continuously for DebounceTime (PUB001)
 *   - Retention:    Held TRUE while VISCOSITY_OK remains TRUE
 *   - Reset:        Immediate on VISCOSITY_OK = FALSE OR PASTE_E_STOP_NC = FALSE (PUB002)
 *   - Same-scan:    Timer PT uses DebounceTime; TON.Q is elapsed >= PT
 *   - Units:        TIME (DebounceTime); TON.ET saturates at PT
 * =============================================================================
 *)
(* CONTRACT_RULES [] *)

    // E-stop immediately clears VFD_RUN and any incomplete debounce state
    IF NOT PASTE_E_STOP_NC THEN
        viscosityValid := FALSE;
        viscosityTimer(IN := FALSE);
        VFD_RUN := FALSE;
    ELSE
        // VISCOSITY_OK must be TRUE for DebounceTime before considered valid
        IF VISCOSITY_OK THEN
            viscosityTimer(IN := TRUE, PT := DebounceTime);
            viscosityValid := viscosityTimer.Q;
        ELSE
            // Immediately invalidate when input becomes FALSE
            viscosityTimer(IN := FALSE);
            viscosityValid := FALSE;
        END_IF;

        // VFD_RUN permitted only when E-stop is safe and viscosity condition is valid
        VFD_RUN := viscosityValid;
    END_IF;

    // Accumulate runtime while VFD_RUN is TRUE
    IF VFD_RUN THEN
        PUMP_RUNTIME_ACC := PUMP_RUNTIME_ACC + TO_LTIME(CycleTime);
    END_IF;

    // Set maintenance indication when threshold reached (informational only)
    IF PUMP_RUNTIME_ACC >= LTIME#500h THEN
        PUMP_MAINT_DUE := TRUE;
    END_IF;

END_FUNCTION_BLOCK

(* ---- public-easy-04.raw_candidate_01.st ---- *)
FUNCTION_BLOCK JamPumpControl
VAR_INPUT
    VISCOSITY_OK    : BOOL;
    PASTE_E_STOP_NC : BOOL;
    DebounceTime    : TIME;
    CycleTime       : TIME;
END_VAR

VAR_OUTPUT
    VFD_RUN          : BOOL := FALSE;
    PUMP_MAINT_DUE   : BOOL := FALSE;
    PUMP_RUNTIME_ACC : LTIME := LTIME#0s;
END_VAR

VAR
    viscosityTimer : TON;
    viscosityValid : BOOL := FALSE;
END_VAR

(* ENGINEERING_CONTRACT
 * =============================================================================
 * Output: VFD_RUN
 *   - Activation:   PASTE_E_STOP_NC = TRUE AND viscosityValid = TRUE (PUB001, PUB002)
 *   - Retention:    Held TRUE while both permissive conditions remain TRUE
 *   - Reset:        Immediate on PASTE_E_STOP_NC = FALSE (E-stop) OR viscosityValid = FALSE
 *   - Same-scan:    E-stop has highest priority; cleared first scan of E-stop event
 *   - Units:        Boolean command, no time units
 * ----------------------------------------------------------------------------
 * Output: PUMP_RUNTIME_ACC
 *   - Activation:   VFD_RUN = TRUE (PUB003)
 *   - Retention:    Preserved while VFD_RUN = FALSE; never cleared by E-stop
 *   - Reset:        None (informational only)
 *   - Same-scan:    Accumulates once per invocation using CycleTime value
 *   - Units:        LTIME nanoseconds; 500h = 1,800,000,000,000 ns (PUB004)
 * ----------------------------------------------------------------------------
 * Output: PUMP_MAINT_DUE
 *   - Activation:   PUMP_RUNTIME_ACC >= 500 hours (PUB004)
 *   - Retention:    Held TRUE once threshold reached (no explicit reset required)
 *   - Reset:        None stated; informational only
 *   - Same-scan:    Evaluated every invocation
 *   - Units:        Boolean indication, does not affect VFD_RUN or safety permissive
 * ----------------------------------------------------------------------------
 * Internal: viscosityValid
 *   - Activation:   VISCOSITY_OK = TRUE continuously for DebounceTime (PUB001)
 *   - Retention:    Held TRUE while VISCOSITY_OK remains TRUE
 *   - Reset:        Immediate on VISCOSITY_OK = FALSE OR PASTE_E_STOP_NC = FALSE (PUB002)
 *   - Same-scan:    Timer PT uses DebounceTime; TON.Q is elapsed >= PT
 *   - Units:        TIME (DebounceTime); TON.ET saturates at PT
 * =============================================================================
 *)
(* CONTRACT_RULES [] *)

    // E-stop immediately clears VFD_RUN and any incomplete debounce state
    IF NOT PASTE_E_STOP_NC THEN
        viscosityValid := FALSE;
        viscosityTimer(IN := FALSE);
        VFD_RUN := FALSE;
    ELSE
        // VISCOSITY_OK must be TRUE for DebounceTime before considered valid
        IF VISCOSITY_OK THEN
            viscosityTimer(IN := TRUE, PT := DebounceTime);
            viscosityValid := viscosityTimer.Q;
        ELSE
            // Immediately invalidate when input becomes FALSE
            viscosityTimer(IN := FALSE);
            viscosityValid := FALSE;
        END_IF;

        // VFD_RUN permitted only when E-stop is safe and viscosity condition is valid
        VFD_RUN := viscosityValid;
    END_IF;

    // Accumulate runtime while VFD_RUN is TRUE
    IF VFD_RUN THEN
        PUMP_RUNTIME_ACC := PUMP_RUNTIME_ACC + TO_LTIME(CycleTime);
    END_IF;

    // Set maintenance indication when threshold reached (informational only)
    IF PUMP_RUNTIME_ACC >= LTIME#500h THEN
        PUMP_MAINT_DUE := TRUE;
    END_IF;

END_FUNCTION_BLOCK

(* ---- public-easy-05.candidate_01.st ---- *)
(* ENGINEERING_CONTRACT *)
(*
  Init period (5s post power-up):
    - PUB001: Operator_Alert=FALSE, Weld_Soft_Start_Active=TRUE, debounce suspended
  Normal monitoring (after init):
    - PUB002: Operator_Alert latches TRUE after Gap_Exceeded TRUE for DebounceTime
    - PUB002: Operator_Alert FALSE immediately when Gap_Exceeded FALSE (alarm clears)
  E-Stop priority:
    - PUB003: Operator_Alert=FALSE immediately, debounce cleared when Weld_E_Stop_NC=FALSE
  Weld_Soft_Start_Active:
    - PUB004: TRUE during init period only; FALSE during normal monitoring and E-Stop
  Timing:
    - PUB005: Init inhibition fixed at 5s (LTIME); DebounceTime must be positive
  Priority hierarchy:
    - PUB006: E-Stop (Weld_E_Stop_NC=FALSE) overrides init and monitoring unconditionally
*)

(* CONTRACT_RULES [{"kind":"hold_until_reset","output":"Operator_Alert","set_input":"Gap_Exceeded","reset_input":"Weld_E_Stop_NC"}] *)

FUNCTION_BLOCK Weld_Gap_Alarm
VAR_INPUT
    Gap_Exceeded : BOOL;
    Weld_E_Stop_NC : BOOL;
    DebounceTime : TIME;
END_VAR
VAR_OUTPUT
    Operator_Alert : BOOL;
    Weld_Soft_Start_Active : BOOL;
END_VAR
VAR
    init_timer : TON;
    debounce_timer : TON;
    tmp_init_done : BOOL;
END_VAR

// E-Stop priority: overrides init and monitoring
IF NOT Weld_E_Stop_NC THEN
    Operator_Alert := FALSE;
    Weld_Soft_Start_Active := FALSE;
    debounce_timer(IN := FALSE, PT := DebounceTime);
    init_timer(IN := FALSE, PT := T#5s);
    tmp_init_done := FALSE;
    RETURN;
END_IF;

// Initialization period (5 seconds)
init_timer(IN := NOT init_timer.Q, PT := T#5s);
Weld_Soft_Start_Active := NOT init_timer.Q;

IF NOT init_timer.Q THEN
    // During initialization: clear debounce
    debounce_timer(IN := FALSE, PT := DebounceTime);
    Operator_Alert := FALSE;
    RETURN;
END_IF;

// Normal monitoring after init complete
tmp_init_done := init_timer.Q;

debounce_timer(IN := Gap_Exceeded AND NOT Operator_Alert, PT := DebounceTime);

IF debounce_timer.Q THEN
    Operator_Alert := TRUE;
ELSIF NOT Gap_Exceeded THEN
    Operator_Alert := FALSE;
END_IF;

END_FUNCTION_BLOCK

(* ---- public-easy-05.raw_candidate_01.st ---- *)
(* ENGINEERING_CONTRACT *)
(*
  Init period (5s post power-up):
    - PUB001: Operator_Alert=FALSE, Weld_Soft_Start_Active=TRUE, debounce suspended
  Normal monitoring (after init):
    - PUB002: Operator_Alert latches TRUE after Gap_Exceeded TRUE for DebounceTime
    - PUB002: Operator_Alert FALSE immediately when Gap_Exceeded FALSE (alarm clears)
  E-Stop priority:
    - PUB003: Operator_Alert=FALSE immediately, debounce cleared when Weld_E_Stop_NC=FALSE
  Weld_Soft_Start_Active:
    - PUB004: TRUE during init period only; FALSE during normal monitoring and E-Stop
  Timing:
    - PUB005: Init inhibition fixed at 5s (LTIME); DebounceTime must be positive
  Priority hierarchy:
    - PUB006: E-Stop (Weld_E_Stop_NC=FALSE) overrides init and monitoring unconditionally
*)

(* CONTRACT_RULES [{"kind":"hold_until_reset","output":"Operator_Alert","set_input":"Gap_Exceeded","reset_input":"Weld_E_Stop_NC"}] *)

FUNCTION_BLOCK Weld_Gap_Alarm
VAR_INPUT
    Gap_Exceeded : BOOL;
    Weld_E_Stop_NC : BOOL;
    DebounceTime : TIME;
END_VAR
VAR_OUTPUT
    Operator_Alert : BOOL;
    Weld_Soft_Start_Active : BOOL;
END_VAR
VAR
    init_timer : TON;
    debounce_timer : TON;
    tmp_init_done : BOOL;
END_VAR

// E-Stop priority: overrides init and monitoring
IF NOT Weld_E_Stop_NC THEN
    Operator_Alert := FALSE;
    Weld_Soft_Start_Active := FALSE;
    debounce_timer(IN := FALSE, PT := DebounceTime);
    init_timer(IN := FALSE, PT := T#5s);
    tmp_init_done := FALSE;
    RETURN;
END_IF;

// Initialization period (5 seconds)
init_timer(IN := NOT init_timer.Q, PT := T#5s);
Weld_Soft_Start_Active := NOT init_timer.Q;

IF NOT init_timer.Q THEN
    // During initialization: clear debounce
    debounce_timer(IN := FALSE, PT := DebounceTime);
    Operator_Alert := FALSE;
    RETURN;
END_IF;

// Normal monitoring after init complete
tmp_init_done := init_timer.Q;

debounce_timer(IN := Gap_Exceeded AND NOT Operator_Alert, PT := DebounceTime);

IF debounce_timer.Q THEN
    Operator_Alert := TRUE;
ELSIF NOT Gap_Exceeded THEN
    Operator_Alert := FALSE;
END_IF;

END_FUNCTION_BLOCK

(* ---- public-easy-06.candidate_01.st ---- *)
(* ENGINEERING_CONTRACT
===================
PUB001: Start demand = DO_LOW AND AERATION_E_STOP_NC (both TRUE required)
PUB002: 5-second PT TON delay; timer enabled while demand active; no edge trigger
PUB003: Immediate BLOWER_RUN disable on demand loss; full 5s delay on re-demand
PUB004: Rising-edge BLOWER_RUN (R_TRIG) increments AERATION_BLOWER_CYCLE_COUNT
PUB005: Power-up initialization: BLOWER_RUN=FALSE, count=0, timer reset

Output state:
- BLOWER_RUN: activation (TON.Q), retention (none - demand-gated),
  explicit reset (demand loss), same-scan priority (timer evaluated each call)
- AERATION_BLOWER_CYCLE_COUNT: increment on BLOWER_RUN rising edge only
*)

(* CONTRACT_RULES [] *)

FUNCTION_BLOCK AerationBlowerControl
VAR_INPUT
    DO_LOW : BOOL;
    AERATION_E_STOP_NC : BOOL;
END_VAR

VAR_OUTPUT
    BLOWER_RUN : BOOL;
    AERATION_BLOWER_CYCLE_COUNT : UINT;
END_VAR

VAR
    StartTimer : TON;
    RunRisingEdge : R_TRIG;
    tmp_DemandActive : BOOL;
END_VAR

// Combine start conditions: DO sufficient AND E-stop inactive
tmp_DemandActive := DO_LOW AND AERATION_E_STOP_NC;

// Rising edge detection for cycle counting
RunRisingEdge(CLK := BLOWER_RUN);

// Increment cycle count on rising edge of BLOWER_RUN
IF RunRisingEdge.Q THEN
    AERATION_BLOWER_CYCLE_COUNT := AERATION_BLOWER_CYCLE_COUNT + UINT#1;
END_IF;

// Timer enabled while demand active
StartTimer(IN := tmp_DemandActive, PT := T#5S);

// Blower control: demand active AND timer elapsed
IF tmp_DemandActive AND StartTimer.Q THEN
    BLOWER_RUN := TRUE;
ELSE
    BLOWER_RUN := FALSE;
END_IF;

END_FUNCTION_BLOCK

(* ---- public-easy-06.patch_base_02.st ---- *)
(* ENGINEERING_CONTRACT
===================
PUB001: Start demand = DO_LOW AND AERATION_E_STOP_NC (both TRUE required)
PUB002: 5-second PT TON delay; timer enabled while demand active; no edge trigger
PUB003: Immediate BLOWER_RUN disable on demand loss; full 5s delay on re-demand
PUB004: Rising-edge BLOWER_RUN (R_TRIG) increments AERATION_BLOWER_CYCLE_COUNT
PUB005: Power-up initialization: BLOWER_RUN=FALSE, count=0, timer reset

Output state:
- BLOWER_RUN: activation (TON.Q), retention (none - demand-gated),
  explicit reset (demand loss), same-scan priority (timer evaluated each call)
- AERATION_BLOWER_CYCLE_COUNT: increment on BLOWER_RUN rising edge only
*)

(* CONTRACT_RULES [] *)

FUNCTION_BLOCK AerationBlowerControl
VAR_INPUT
    DO_LOW : BOOL;
    AERATION_E_STOP_NC : BOOL;
END_VAR

VAR_OUTPUT
    BLOWER_RUN : BOOL;
    AERATION_BLOWER_CYCLE_COUNT : UINT;
END_VAR

VAR
    StartTimer : TON;
    RunRisingEdge : R_TRIG;
    tmp_DemandActive : BOOL;
END_VAR

// Combine start conditions: DO sufficient AND E-stop inactive
tmp_DemandActive := DO_LOW AND AERATION_E_STOP_NC;

// Rising edge detection for cycle counting
RunRisingEdge(CLK := BLOWER_RUN);

// Increment cycle count on rising edge of BLOWER_RUN
IF RunRisingEdge.Q THEN
    AERATION_BLOWER_CYCLE_COUNT := AERATION_BLOWER_CYCLE_COUNT + UINT#1;
END_IF;

// Timer enabled while demand active
StartTimer(IN := tmp_DemandActive, PT := T#5S);

// Blower control: demand active AND timer elapsed
IF tmp_DemandActive AND StartTimer.Q THEN
    BLOWER_RUN := TRUE;
ELSE
    BLOWER_RUN := FALSE;
END_IF;

END_FUNCTION_BLOCK

(* ---- public-easy-06.raw_candidate_01.st ---- *)
(* ENGINEERING_CONTRACT
===================
PUB001: Start demand = DO_LOW AND AERATION_E_STOP_NC (both TRUE required)
PUB002: 5-second PT TON delay; timer enabled while demand active; no edge trigger
PUB003: Immediate BLOWER_RUN disable on demand loss; full 5s delay on re-demand
PUB004: Rising-edge BLOWER_RUN (R_TRIG) increments AERATION_BLOWER_CYCLE_COUNT
PUB005: Power-up initialization: BLOWER_RUN=FALSE, count=0, timer reset

Output state:
- BLOWER_RUN: activation (TON.Q), retention (none - demand-gated),
  explicit reset (demand loss), same-scan priority (timer evaluated each call)
- AERATION_BLOWER_CYCLE_COUNT: increment on BLOWER_RUN rising edge only
*)

(* CONTRACT_RULES [] *)

FUNCTION_BLOCK AerationBlowerControl
VAR_INPUT
    DO_LOW : BOOL;
    AERATION_E_STOP_NC : BOOL;
END_VAR

VAR_OUTPUT
    BLOWER_RUN : BOOL;
    AERATION_BLOWER_CYCLE_COUNT : UINT;
END_VAR

VAR
    StartTimer : TON;
    RunRisingEdge : R_TRIG;
    tmp_DemandActive : BOOL;
END_VAR

// Combine start conditions: DO sufficient AND E-stop inactive
tmp_DemandActive := DO_LOW AND AERATION_E_STOP_NC;

// Rising edge detection for cycle counting
RunRisingEdge(CLK := BLOWER_RUN);

// Increment cycle count on rising edge of BLOWER_RUN
IF RunRisingEdge.Q THEN
    AERATION_BLOWER_CYCLE_COUNT := AERATION_BLOWER_CYCLE_COUNT + UINT#1;
END_IF;

// Timer enabled while demand active
StartTimer(IN := tmp_DemandActive, PT := T#5S);

// Blower control: demand active AND timer elapsed
IF tmp_DemandActive AND StartTimer.Q THEN
    BLOWER_RUN := TRUE;
ELSE
    BLOWER_RUN := FALSE;
END_IF;

END_FUNCTION_BLOCK

(* ---- public-hard-01.candidate_01.st ---- *)
FUNCTION_BLOCK MaterialProportioning
VAR_INPUT
    estop           : BOOL;          // Emergency stop signal (FALSE = stopped)
    opeMode         : BOOL;          // Operation mode (FALSE = manual, TRUE = automatic)
    valveAStart     : BOOL;          // Valve A start button
    valveBStart     : BOOL;          // Valve B start button
    valveCStart     : BOOL;          // Valve C start button
    valveDStart     : BOOL;          // Valve D start button
    mixMotorStart   : BOOL;          // Mixing motor start button
    autoStart       : BOOL;          // Automatic start button
    processMode     : BOOL;          // Process mode (FALSE = simple, TRUE = with C)
    levelSensor     : INT;           // Liquid level sensor (cm)
    mixMotorComplete: BOOL;          // Mixing complete signal
END_VAR
VAR_OUTPUT
    valveARun       : BOOL;          // Valve A run command
    valveBRun       : BOOL;          // Valve B run command
    valveCRun       : BOOL;          // Valve C run command
    valveDRun       : BOOL;          // Valve D run command
    mixMotorRun     : BOOL;          // Mixing motor run command
END_VAR
VAR
    // Rising edge detection for manual toggle buttons
    tmp_autoStart rising  : R_TRIG;
    tmp_valveAStart rising: R_TRIG;
    tmp_valveBStart rising: R_TRIG;
    tmp_valveCStart rising: R_TRIG;
    tmp_valveDStart rising: R_TRIG;
    tmp_mixMotorStart rising: R_TRIG;

    // Automatic mode state machine
    tmp_autoState   : INT;           // 0=idle, 1=fillA, 2=fillB, 3=fillC, 4=mix, 5=drain, 6=done

    // Manual mode toggle states
    tmp_manualValveA    : BOOL;
    tmp_manualValveB    : BOOL;
    tmp_manualValveC    : BOOL;
    tmp_manualValveD    : BOOL;
    tmp_manualMixMotor  : BOOL;

    // Process complete flag for automatic mode
    tmp_autoComplete    : BOOL;
END_VAR

(* ENGINEERING_CONTRACT
================================================================================
Output          | Activation                  | Retention      | Reset
----------------|------------------------------|----------------|-------------------------
valveARun       | Manual: rising valveAStart   | Hold toggle    | estop, opeMode, auto step
                | Auto: state=1, level<50      |                |
PUB001, PUB002, PUB003, PUB004, PUB005, PUB006, PUB007, PUB008
----------------|------------------------------|----------------|-------------------------
valveBRun       | Auto: state=2, level<80      | Hold until 80cm| estop, opeMode, auto step
                |                              |                |
PUB003, PUB004, PUB006, PUB007, PUB008
----------------|------------------------------|----------------|-------------------------
valveCRun       | Auto: state=3, level<100     | Hold until 100cm| estop, opeMode, auto step
                | (processMode=true only)      |                |
PUB003, PUB004, PUB006, PUB007, PUB008
----------------|------------------------------|----------------|-------------------------
valveDRun       | Auto: mixMotorComplete       | Hold until reset| estop, opeMode, autoStart
                |                              |                |
PUB007, PUB008, PUB011, PUB012, PUB013, PUB014, PUB015
----------------|------------------------------|----------------|-------------------------
mixMotorRun     | Auto: state=4                | Hold until complete| estop, opeMode, autoStart
                | Manual: rising mixMotorStart |                |
PUB007, PUB008, PUB011, PUB012, PUB013, PUB014, PUB015
================================================================================
Priority: estop > manual/automatic mode switch > same-scan state updates
Boundary: levelSensor thresholds at 50cm, 80cm, 100cm (>= comparisons)
================================================================================
*)

(* CONTRACT_RULES [] *)

// Detect rising edges for toggle buttons
rising(autoStart);
rising(valveAStart);
rising(valveBStart);
rising(valveCStart);
rising(valveDStart);
rising(mixMotorStart);

// Emergency stop: all equipment OFF immediately
IF NOT estop THEN
    valveARun := FALSE;
    valveBRun := FALSE;
    valveCRun := FALSE;
    valveDRun := FALSE;
    mixMotorRun := FALSE;
    tmp_autoState := 0;
    tmp_autoComplete := FALSE;
    tmp_manualValveA := FALSE;
    tmp_manualValveB := FALSE;
    tmp_manualValveC := FALSE;
    tmp_manualValveD := FALSE;
    tmp_manualMixMotor := FALSE;
    RETURN;
END_IF;

// Mode selection
IF opeMode THEN
    // AUTOMATIC MODE
    // Rising edge of autoStart initiates process
    IF rising.Q AND tmp_autoState = 0 THEN
        tmp_autoState := 1;
        tmp_autoComplete := FALSE;
    END_IF;

    // State machine execution
    CASE tmp_autoState OF
        0:  // Idle - all off
            valveARun := FALSE;
            valveBRun := FALSE;
            valveCRun := FALSE;
            valveDRun := FALSE;
            mixMotorRun := FALSE;

        1:  // Fill with valve A until level >= 50cm
            valveARun := TRUE;
            valveBRun := FALSE;
            valveCRun := FALSE;
            valveDRun := FALSE;
            mixMotorRun := FALSE;
            IF levelSensor >= 50 THEN
                valveARun := FALSE;
                tmp_autoState := 2;
            END_IF;

        2:  // Fill with valve B until level >= 80cm
            valveARun := FALSE;
            valveBRun := TRUE;
            valveCRun := FALSE;
            valveDRun := FALSE;
            mixMotorRun := FALSE;
            IF levelSensor >= 80 THEN
                valveBRun := FALSE;
                // Check processMode to determine next state
                IF processMode THEN
                    tmp_autoState := 3;  // Go to valve C
                ELSE
                    tmp_autoState := 4;  // Go directly to mixing
                END_IF;
            END_IF;

        3:  // Fill with valve C (processMode=true) until level >= 100cm
            valveARun := FALSE;
            valveBRun := FALSE;
            valveCRun := TRUE;
            valveDRun := FALSE;
            mixMotorRun := FALSE;
            IF levelSensor >= 100 THEN
                valveCRun := FALSE;
                tmp_autoState := 4;
            END_IF;

        4:  // Mixing until mixMotorComplete signal
            valveARun := FALSE;
            valveBRun := FALSE;
            valveCRun := FALSE;
            valveDRun := FALSE;
            mixMotorRun := TRUE;
            IF mixMotorComplete THEN
                mixMotorRun := FALSE;
                tmp_autoState := 5;
            END_IF;

        5:  // Open valve D to drain
            valveARun := FALSE;
            valveBRun := FALSE;
            valveCRun := FALSE;
            valveDRun := TRUE;
            mixMotorRun := FALSE;
            tmp_autoComplete := TRUE;
            tmp_autoState := 6;

        6:  // Process complete - valve D remains open until reset
            valveARun := FALSE;
            valveBRun := FALSE;
            valveCRun := FALSE;
            valveDRun := TRUE;
            mixMotorRun := FALSE;
            // Wait for autoStart to reset
            IF rising.Q THEN
                tmp_autoState := 0;
                tmp_autoComplete := FALSE;
            END_IF;
    END_CASE;

ELSE
    // MANUAL MODE
    // Reset automatic state when switching to manual
    tmp_autoState := 0;
    tmp_autoComplete := FALSE;

    // Toggle valve A
    IF rising(valveAStart) THEN
        tmp_manualValveA := NOT tmp_manualValveA;
    END_IF;

    // Toggle valve B
    IF rising(valveBStart) THEN
        tmp_manualValveB := NOT tmp_manualValveB;
    END_IF;

    // Toggle valve C
    IF rising(valveCStart) THEN
        tmp_manualValveC := NOT tmp_manualValveC;
    END_IF;

    // Toggle valve D
    IF rising(valveDStart) THEN
        tmp_manualValveD := NOT tmp_manualValveD;
    END_IF;

    // Toggle mixing motor
    IF rising(mixMotorStart) THEN
        tmp_manualMixMotor := NOT tmp_manualMixMotor;
    END_IF;

    // Assign manual toggle states to outputs
    valveARun := tmp_manualValveA;
    valveBRun := tmp_manualValveB;
    valveCRun := tmp_manualValveC;
    valveDRun := tmp_manualValveD;
    mixMotorRun := tmp_manualMixMotor;
END_IF;

END_FUNCTION_BLOCK

(* ---- public-hard-01.candidate_02.st ---- *)
FUNCTION_BLOCK MaterialProportioning
VAR_INPUT
    estop           : BOOL;          // Emergency stop signal (FALSE = stopped)
    opeMode         : BOOL;          // Operation mode (FALSE = manual, TRUE = automatic)
    valveAStart     : BOOL;          // Valve A start button
    valveBStart     : BOOL;          // Valve B start button
    valveCStart     : BOOL;          // Valve C start button
    valveDStart     : BOOL;          // Valve D start button
    mixMotorStart   : BOOL;          // Mixing motor start button
    autoStart       : BOOL;          // Automatic start button
    processMode     : BOOL;          // Process mode (FALSE = simple, TRUE = with C)
    levelSensor     : INT;           // Liquid level sensor (cm)
    mixMotorComplete: BOOL;          // Mixing complete signal
END_VAR
VAR_OUTPUT
    valveARun       : BOOL;          // Valve A run command
    valveBRun       : BOOL;          // Valve B run command
    valveCRun       : BOOL;          // Valve C run command
    valveDRun       : BOOL;          // Valve D run command
    mixMotorRun     : BOOL;          // Mixing motor run command
END_VAR
VAR
    // Rising edge detection for manual toggle buttons
    tmp_autoStart        : R_TRIG;
    tmp_valveAStart      : R_TRIG;
    tmp_valveBStart      : R_TRIG;
    tmp_valveCStart      : R_TRIG;
    tmp_valveDStart      : R_TRIG;
    tmp_mixMotorStart    : R_TRIG;

    // Automatic mode state machine
    tmp_autoState   : INT;           // 0=idle, 1=fillA, 2=fillB, 3=fillC, 4=mix, 5=drain, 6=done

    // Manual mode toggle states
    tmp_manualValveA    : BOOL;
    tmp_manualValveB    : BOOL;
    tmp_manualValveC    : BOOL;
    tmp_manualValveD    : BOOL;
    tmp_manualMixMotor  : BOOL;

    // Process complete flag for automatic mode
    tmp_autoComplete    : BOOL;
END_VAR

(* ENGINEERING_CONTRACT
================================================================================
Output          | Activation                  | Retention      | Reset
----------------|------------------------------|----------------|-------------------------
valveARun       | Manual: rising valveAStart   | Hold toggle    | estop, opeMode, auto step
                | Auto: state=1, level<50      |                |
PUB001, PUB002, PUB003, PUB004, PUB005, PUB006, PUB007, PUB008
----------------|------------------------------|----------------|-------------------------
valveBRun       | Auto: state=2, level<80      | Hold until 80cm| estop, opeMode, auto step
                |                              |                |
PUB003, PUB004, PUB006, PUB007, PUB008
----------------|------------------------------|----------------|-------------------------
valveCRun       | Auto: state=3, level<100     | Hold until 100cm| estop, opeMode, auto step
                | (processMode=true only)      |                |
PUB003, PUB004, PUB006, PUB007, PUB008
----------------|------------------------------|----------------|-------------------------
valveDRun       | Auto: mixMotorComplete       | Hold until reset| estop, opeMode, autoStart
                |                              |                |
PUB007, PUB008, PUB011, PUB012, PUB013, PUB014, PUB015
----------------|------------------------------|----------------|-------------------------
mixMotorRun     | Auto: state=4                | Hold until complete| estop, opeMode, autoStart
                | Manual: rising mixMotorStart |                |
PUB007, PUB008, PUB011, PUB012, PUB013, PUB014, PUB015
================================================================================
Priority: estop > manual/automatic mode switch > same-scan state updates
Boundary: levelSensor thresholds at 50cm, 80cm, 100cm (>= comparisons)
================================================================================
*)

(* CONTRACT_RULES [] *)

// Detect rising edges for toggle buttons
tmp_autoStart(CLK := autoStart);
tmp_valveAStart(CLK := valveAStart);
tmp_valveBStart(CLK := valveBStart);
tmp_valveCStart(CLK := valveCStart);
tmp_valveDStart(CLK := valveDStart);
tmp_mixMotorStart(CLK := mixMotorStart);

// Emergency stop: all equipment OFF immediately
IF NOT estop THEN
    valveARun := FALSE;
    valveBRun := FALSE;
    valveCRun := FALSE;
    valveDRun := FALSE;
    mixMotorRun := FALSE;
    tmp_autoState := 0;
    tmp_autoComplete := FALSE;
    tmp_manualValveA := FALSE;
    tmp_manualValveB := FALSE;
    tmp_manualValveC := FALSE;
    tmp_manualValveD := FALSE;
    tmp_manualMixMotor := FALSE;
    RETURN;
END_IF;

// Mode selection
IF opeMode THEN
    // AUTOMATIC MODE
    // Rising edge of autoStart initiates process
    IF tmp_autoStart.Q AND tmp_autoState = 0 THEN
        tmp_autoState := 1;
        tmp_autoComplete := FALSE;
    END_IF;

    // State machine execution
    CASE tmp_autoState OF
        0:  // Idle - all off
            valveARun := FALSE;
            valveBRun := FALSE;
            valveCRun := FALSE;
            valveDRun := FALSE;
            mixMotorRun := FALSE;

        1:  // Fill with valve A until level >= 50cm
            valveARun := TRUE;
            valveBRun := FALSE;
            valveCRun := FALSE;
            valveDRun := FALSE;
            mixMotorRun := FALSE;
            IF levelSensor >= 50 THEN
                valveARun := FALSE;
                tmp_autoState := 2;
            END_IF;

        2:  // Fill with valve B until level >= 80cm
            valveARun := FALSE;
            valveBRun := TRUE;
            valveCRun := FALSE;
            valveDRun := FALSE;
            mixMotorRun := FALSE;
            IF levelSensor >= 80 THEN
                valveBRun := FALSE;
                // Check processMode to determine next state
                IF processMode THEN
                    tmp_autoState := 3;  // Go to valve C
                ELSE
                    tmp_autoState := 4;  // Go directly to mixing
                END_IF;
            END_IF;

        3:  // Fill with valve C (processMode=true) until level >= 100cm
            valveARun := FALSE;
            valveBRun := FALSE;
            valveCRun := TRUE;
            valveDRun := FALSE;
            mixMotorRun := FALSE;
            IF levelSensor >= 100 THEN
                valveCRun := FALSE;
                tmp_autoState := 4;
            END_IF;

        4:  // Mixing until mixMotorComplete signal
            valveARun := FALSE;
            valveBRun := FALSE;
            valveCRun := FALSE;
            valveDRun := FALSE;
            mixMotorRun := TRUE;
            IF mixMotorComplete THEN
                mixMotorRun := FALSE;
                tmp_autoState := 5;
            END_IF;

        5:  // Open valve D to drain
            valveARun := FALSE;
            valveBRun := FALSE;
            valveCRun := FALSE;
            valveDRun := TRUE;
            mixMotorRun := FALSE;
            tmp_autoComplete := TRUE;
            tmp_autoState := 6;

        6:  // Process complete - valve D remains open until reset
            valveARun := FALSE;
            valveBRun := FALSE;
            valveCRun := FALSE;
            valveDRun := TRUE;
            mixMotorRun := FALSE;
            // Wait for autoStart to reset
            IF tmp_autoStart.Q THEN
                tmp_autoState := 0;
                tmp_autoComplete := FALSE;
            END_IF;
    END_CASE;

ELSE
    // MANUAL MODE
    // Reset automatic state when switching to manual
    tmp_autoState := 0;
    tmp_autoComplete := FALSE;

    // Toggle valve A
    IF tmp_valveAStart.Q THEN
        tmp_manualValveA := NOT tmp_manualValveA;
    END_IF;

    // Toggle valve B
    IF tmp_valveBStart.Q THEN
        tmp_manualValveB := NOT tmp_manualValveB;
    END_IF;

    // Toggle valve C
    IF tmp_valveCStart.Q THEN
        tmp_manualValveC := NOT tmp_manualValveC;
    END_IF;

    // Toggle valve D
    IF tmp_valveDStart.Q THEN
        tmp_manualValveD := NOT tmp_manualValveD;
    END_IF;

    // Toggle mixing motor
    IF tmp_mixMotorStart.Q THEN
        tmp_manualMixMotor := NOT tmp_manualMixMotor;
    END_IF;

    // Assign manual toggle states to outputs
    valveARun := tmp_manualValveA;
    valveBRun := tmp_manualValveB;
    valveCRun := tmp_manualValveC;
    valveDRun := tmp_manualValveD;
    mixMotorRun := tmp_manualMixMotor;
END_IF;

END_FUNCTION_BLOCK

(* ---- public-hard-01.patch_base_02.st ---- *)
FUNCTION_BLOCK MaterialProportioning
VAR_INPUT
    estop           : BOOL;          // Emergency stop signal (FALSE = stopped)
    opeMode         : BOOL;          // Operation mode (FALSE = manual, TRUE = automatic)
    valveAStart     : BOOL;          // Valve A start button
    valveBStart     : BOOL;          // Valve B start button
    valveCStart     : BOOL;          // Valve C start button
    valveDStart     : BOOL;          // Valve D start button
    mixMotorStart   : BOOL;          // Mixing motor start button
    autoStart       : BOOL;          // Automatic start button
    processMode     : BOOL;          // Process mode (FALSE = simple, TRUE = with C)
    levelSensor     : INT;           // Liquid level sensor (cm)
    mixMotorComplete: BOOL;          // Mixing complete signal
END_VAR
VAR_OUTPUT
    valveARun       : BOOL;          // Valve A run command
    valveBRun       : BOOL;          // Valve B run command
    valveCRun       : BOOL;          // Valve C run command
    valveDRun       : BOOL;          // Valve D run command
    mixMotorRun     : BOOL;          // Mixing motor run command
END_VAR
VAR
    // Rising edge detection for manual toggle buttons
    tmp_autoStart rising  : R_TRIG;
    tmp_valveAStart rising: R_TRIG;
    tmp_valveBStart rising: R_TRIG;
    tmp_valveCStart rising: R_TRIG;
    tmp_valveDStart rising: R_TRIG;
    tmp_mixMotorStart rising: R_TRIG;

    // Automatic mode state machine
    tmp_autoState   : INT;           // 0=idle, 1=fillA, 2=fillB, 3=fillC, 4=mix, 5=drain, 6=done

    // Manual mode toggle states
    tmp_manualValveA    : BOOL;
    tmp_manualValveB    : BOOL;
    tmp_manualValveC    : BOOL;
    tmp_manualValveD    : BOOL;
    tmp_manualMixMotor  : BOOL;

    // Process complete flag for automatic mode
    tmp_autoComplete    : BOOL;
END_VAR

(* ENGINEERING_CONTRACT
================================================================================
Output          | Activation                  | Retention      | Reset
----------------|------------------------------|----------------|-------------------------
valveARun       | Manual: rising valveAStart   | Hold toggle    | estop, opeMode, auto step
                | Auto: state=1, level<50      |                |
PUB001, PUB002, PUB003, PUB004, PUB005, PUB006, PUB007, PUB008
----------------|------------------------------|----------------|-------------------------
valveBRun       | Auto: state=2, level<80      | Hold until 80cm| estop, opeMode, auto step
                |                              |                |
PUB003, PUB004, PUB006, PUB007, PUB008
----------------|------------------------------|----------------|-------------------------
valveCRun       | Auto: state=3, level<100     | Hold until 100cm| estop, opeMode, auto step
                | (processMode=true only)      |                |
PUB003, PUB004, PUB006, PUB007, PUB008
----------------|------------------------------|----------------|-------------------------
valveDRun       | Auto: mixMotorComplete       | Hold until reset| estop, opeMode, autoStart
                |                              |                |
PUB007, PUB008, PUB011, PUB012, PUB013, PUB014, PUB015
----------------|------------------------------|----------------|-------------------------
mixMotorRun     | Auto: state=4                | Hold until complete| estop, opeMode, autoStart
                | Manual: rising mixMotorStart |                |
PUB007, PUB008, PUB011, PUB012, PUB013, PUB014, PUB015
================================================================================
Priority: estop > manual/automatic mode switch > same-scan state updates
Boundary: levelSensor thresholds at 50cm, 80cm, 100cm (>= comparisons)
================================================================================
*)

(* CONTRACT_RULES [] *)

// Detect rising edges for toggle buttons
rising(autoStart);
rising(valveAStart);
rising(valveBStart);
rising(valveCStart);
rising(valveDStart);
rising(mixMotorStart);

// Emergency stop: all equipment OFF immediately
IF NOT estop THEN
    valveARun := FALSE;
    valveBRun := FALSE;
    valveCRun := FALSE;
    valveDRun := FALSE;
    mixMotorRun := FALSE;
    tmp_autoState := 0;
    tmp_autoComplete := FALSE;
    tmp_manualValveA := FALSE;
    tmp_manualValveB := FALSE;
    tmp_manualValveC := FALSE;
    tmp_manualValveD := FALSE;
    tmp_manualMixMotor := FALSE;
    RETURN;
END_IF;

// Mode selection
IF opeMode THEN
    // AUTOMATIC MODE
    // Rising edge of autoStart initiates process
    IF rising.Q AND tmp_autoState = 0 THEN
        tmp_autoState := 1;
        tmp_autoComplete := FALSE;
    END_IF;

    // State machine execution
    CASE tmp_autoState OF
        0:  // Idle - all off
            valveARun := FALSE;
            valveBRun := FALSE;
            valveCRun := FALSE;
            valveDRun := FALSE;
            mixMotorRun := FALSE;

        1:  // Fill with valve A until level >= 50cm
            valveARun := TRUE;
            valveBRun := FALSE;
            valveCRun := FALSE;
            valveDRun := FALSE;
            mixMotorRun := FALSE;
            IF levelSensor >= 50 THEN
                valveARun := FALSE;
                tmp_autoState := 2;
            END_IF;

        2:  // Fill with valve B until level >= 80cm
            valveARun := FALSE;
            valveBRun := TRUE;
            valveCRun := FALSE;
            valveDRun := FALSE;
            mixMotorRun := FALSE;
            IF levelSensor >= 80 THEN
                valveBRun := FALSE;
                // Check processMode to determine next state
                IF processMode THEN
                    tmp_autoState := 3;  // Go to valve C
                ELSE
                    tmp_autoState := 4;  // Go directly to mixing
                END_IF;
            END_IF;

        3:  // Fill with valve C (processMode=true) until level >= 100cm
            valveARun := FALSE;
            valveBRun := FALSE;
            valveCRun := TRUE;
            valveDRun := FALSE;
            mixMotorRun := FALSE;
            IF levelSensor >= 100 THEN
                valveCRun := FALSE;
                tmp_autoState := 4;
            END_IF;

        4:  // Mixing until mixMotorComplete signal
            valveARun := FALSE;
            valveBRun := FALSE;
            valveCRun := FALSE;
            valveDRun := FALSE;
            mixMotorRun := TRUE;
            IF mixMotorComplete THEN
                mixMotorRun := FALSE;
                tmp_autoState := 5;
            END_IF;

        5:  // Open valve D to drain
            valveARun := FALSE;
            valveBRun := FALSE;
            valveCRun := FALSE;
            valveDRun := TRUE;
            mixMotorRun := FALSE;
            tmp_autoComplete := TRUE;
            tmp_autoState := 6;

        6:  // Process complete - valve D remains open until reset
            valveARun := FALSE;
            valveBRun := FALSE;
            valveCRun := FALSE;
            valveDRun := TRUE;
            mixMotorRun := FALSE;
            // Wait for autoStart to reset
            IF rising.Q THEN
                tmp_autoState := 0;
                tmp_autoComplete := FALSE;
            END_IF;
    END_CASE;

ELSE
    // MANUAL MODE
    // Reset automatic state when switching to manual
    tmp_autoState := 0;
    tmp_autoComplete := FALSE;

    // Toggle valve A
    IF rising(valveAStart) THEN
        tmp_manualValveA := NOT tmp_manualValveA;
    END_IF;

    // Toggle valve B
    IF rising(valveBStart) THEN
        tmp_manualValveB := NOT tmp_manualValveB;
    END_IF;

    // Toggle valve C
    IF rising(valveCStart) THEN
        tmp_manualValveC := NOT tmp_manualValveC;
    END_IF;

    // Toggle valve D
    IF rising(valveDStart) THEN
        tmp_manualValveD := NOT tmp_manualValveD;
    END_IF;

    // Toggle mixing motor
    IF rising(mixMotorStart) THEN
        tmp_manualMixMotor := NOT tmp_manualMixMotor;
    END_IF;

    // Assign manual toggle states to outputs
    valveARun := tmp_manualValveA;
    valveBRun := tmp_manualValveB;
    valveCRun := tmp_manualValveC;
    valveDRun := tmp_manualValveD;
    mixMotorRun := tmp_manualMixMotor;
END_IF;

END_FUNCTION_BLOCK

(* ---- public-hard-01.raw_candidate_01.st ---- *)
FUNCTION_BLOCK MaterialProportioning
VAR_INPUT
    estop           : BOOL;          // Emergency stop signal (FALSE = stopped)
    opeMode         : BOOL;          // Operation mode (FALSE = manual, TRUE = automatic)
    valveAStart     : BOOL;          // Valve A start button
    valveBStart     : BOOL;          // Valve B start button
    valveCStart     : BOOL;          // Valve C start button
    valveDStart     : BOOL;          // Valve D start button
    mixMotorStart   : BOOL;          // Mixing motor start button
    autoStart       : BOOL;          // Automatic start button
    processMode     : BOOL;          // Process mode (FALSE = simple, TRUE = with C)
    levelSensor     : INT;           // Liquid level sensor (cm)
    mixMotorComplete: BOOL;          // Mixing complete signal
END_VAR
VAR_OUTPUT
    valveARun       : BOOL;          // Valve A run command
    valveBRun       : BOOL;          // Valve B run command
    valveCRun       : BOOL;          // Valve C run command
    valveDRun       : BOOL;          // Valve D run command
    mixMotorRun     : BOOL;          // Mixing motor run command
END_VAR
VAR
    // Rising edge detection for manual toggle buttons
    tmp_autoStart rising  : R_TRIG;
    tmp_valveAStart rising: R_TRIG;
    tmp_valveBStart rising: R_TRIG;
    tmp_valveCStart rising: R_TRIG;
    tmp_valveDStart rising: R_TRIG;
    tmp_mixMotorStart rising: R_TRIG;

    // Automatic mode state machine
    tmp_autoState   : INT;           // 0=idle, 1=fillA, 2=fillB, 3=fillC, 4=mix, 5=drain, 6=done

    // Manual mode toggle states
    tmp_manualValveA    : BOOL;
    tmp_manualValveB    : BOOL;
    tmp_manualValveC    : BOOL;
    tmp_manualValveD    : BOOL;
    tmp_manualMixMotor  : BOOL;

    // Process complete flag for automatic mode
    tmp_autoComplete    : BOOL;
END_VAR

(* ENGINEERING_CONTRACT
================================================================================
Output          | Activation                  | Retention      | Reset
----------------|------------------------------|----------------|-------------------------
valveARun       | Manual: rising valveAStart   | Hold toggle    | estop, opeMode, auto step
                | Auto: state=1, level<50      |                |
PUB001, PUB002, PUB003, PUB004, PUB005, PUB006, PUB007, PUB008
----------------|------------------------------|----------------|-------------------------
valveBRun       | Auto: state=2, level<80      | Hold until 80cm| estop, opeMode, auto step
                |                              |                |
PUB003, PUB004, PUB006, PUB007, PUB008
----------------|------------------------------|----------------|-------------------------
valveCRun       | Auto: state=3, level<100     | Hold until 100cm| estop, opeMode, auto step
                | (processMode=true only)      |                |
PUB003, PUB004, PUB006, PUB007, PUB008
----------------|------------------------------|----------------|-------------------------
valveDRun       | Auto: mixMotorComplete       | Hold until reset| estop, opeMode, autoStart
                |                              |                |
PUB007, PUB008, PUB011, PUB012, PUB013, PUB014, PUB015
----------------|------------------------------|----------------|-------------------------
mixMotorRun     | Auto: state=4                | Hold until complete| estop, opeMode, autoStart
                | Manual: rising mixMotorStart |                |
PUB007, PUB008, PUB011, PUB012, PUB013, PUB014, PUB015
================================================================================
Priority: estop > manual/automatic mode switch > same-scan state updates
Boundary: levelSensor thresholds at 50cm, 80cm, 100cm (>= comparisons)
================================================================================
*)

(* CONTRACT_RULES [] *)

// Detect rising edges for toggle buttons
rising(autoStart);
rising(valveAStart);
rising(valveBStart);
rising(valveCStart);
rising(valveDStart);
rising(mixMotorStart);

// Emergency stop: all equipment OFF immediately
IF NOT estop THEN
    valveARun := FALSE;
    valveBRun := FALSE;
    valveCRun := FALSE;
    valveDRun := FALSE;
    mixMotorRun := FALSE;
    tmp_autoState := 0;
    tmp_autoComplete := FALSE;
    tmp_manualValveA := FALSE;
    tmp_manualValveB := FALSE;
    tmp_manualValveC := FALSE;
    tmp_manualValveD := FALSE;
    tmp_manualMixMotor := FALSE;
    RETURN;
END_IF

// Mode selection
IF opeMode THEN
    // AUTOMATIC MODE
    // Rising edge of autoStart initiates process
    IF rising.Q AND tmp_autoState = 0 THEN
        tmp_autoState := 1;
        tmp_autoComplete := FALSE;
    END_IF

    // State machine execution
    CASE tmp_autoState OF
        0:  // Idle - all off
            valveARun := FALSE;
            valveBRun := FALSE;
            valveCRun := FALSE;
            valveDRun := FALSE;
            mixMotorRun := FALSE;

        1:  // Fill with valve A until level >= 50cm
            valveARun := TRUE;
            valveBRun := FALSE;
            valveCRun := FALSE;
            valveDRun := FALSE;
            mixMotorRun := FALSE;
            IF levelSensor >= 50 THEN
                valveARun := FALSE;
                tmp_autoState := 2;
            END_IF

        2:  // Fill with valve B until level >= 80cm
            valveARun := FALSE;
            valveBRun := TRUE;
            valveCRun := FALSE;
            valveDRun := FALSE;
            mixMotorRun := FALSE;
            IF levelSensor >= 80 THEN
                valveBRun := FALSE;
                // Check processMode to determine next state
                IF processMode THEN
                    tmp_autoState := 3;  // Go to valve C
                ELSE
                    tmp_autoState := 4;  // Go directly to mixing
                END_IF
            END_IF

        3:  // Fill with valve C (processMode=true) until level >= 100cm
            valveARun := FALSE;
            valveBRun := FALSE;
            valveCRun := TRUE;
            valveDRun := FALSE;
            mixMotorRun := FALSE;
            IF levelSensor >= 100 THEN
                valveCRun := FALSE;
                tmp_autoState := 4;
            END_IF

        4:  // Mixing until mixMotorComplete signal
            valveARun := FALSE;
            valveBRun := FALSE;
            valveCRun := FALSE;
            valveDRun := FALSE;
            mixMotorRun := TRUE;
            IF mixMotorComplete THEN
                mixMotorRun := FALSE;
                tmp_autoState := 5;
            END_IF

        5:  // Open valve D to drain
            valveARun := FALSE;
            valveBRun := FALSE;
            valveCRun := FALSE;
            valveDRun := TRUE;
            mixMotorRun := FALSE;
            tmp_autoComplete := TRUE;
            tmp_autoState := 6;

        6:  // Process complete - valve D remains open until reset
            valveARun := FALSE;
            valveBRun := FALSE;
            valveCRun := FALSE;
            valveDRun := TRUE;
            mixMotorRun := FALSE;
            // Wait for autoStart to reset
            IF rising.Q THEN
                tmp_autoState := 0;
                tmp_autoComplete := FALSE;
            END_IF
    END_CASE

ELSE
    // MANUAL MODE
    // Reset automatic state when switching to manual
    tmp_autoState := 0;
    tmp_autoComplete := FALSE;

    // Toggle valve A
    IF rising(valveAStart) THEN
        tmp_manualValveA := NOT tmp_manualValveA;
    END_IF

    // Toggle valve B
    IF rising(valveBStart) THEN
        tmp_manualValveB := NOT tmp_manualValveB;
    END_IF

    // Toggle valve C
    IF rising(valveCStart) THEN
        tmp_manualValveC := NOT tmp_manualValveC;
    END_IF

    // Toggle valve D
    IF rising(valveDStart) THEN
        tmp_manualValveD := NOT tmp_manualValveD;
    END_IF

    // Toggle mixing motor
    IF rising(mixMotorStart) THEN
        tmp_manualMixMotor := NOT tmp_manualMixMotor;
    END_IF

    // Assign manual toggle states to outputs
    valveARun := tmp_manualValveA;
    valveBRun := tmp_manualValveB;
    valveCRun := tmp_manualValveC;
    valveDRun := tmp_manualValveD;
    mixMotorRun := tmp_manualMixMotor;
END_IF

END_FUNCTION_BLOCK
